(* IEC 61131-3 sources: iecf/harness/cases, 218 files *)

(* ---- autoaddrsections.st ---- *)
(* TwinCAT's `*` structures where Ed.3 6.4.4.8 refuses them
   (auto-addresses, W0020), as TcOpen's TcoEthercatMasterDevice: a
   block's VAR_INPUT, placed per instance as a VAR's, and a method's
   VAR, plain memory of the call; and its VAR_OUTPUT, which Ed.3
   allows, placed per instance.
   Placed by path, nothing stated: M: P.M.INPUTS.A 0, P.SRC.A 2.
   Q: P.M.INPUTS.B 0, P.M.OUTPUTS.Q 2, P.SRC.B 4.
   Worked by hand, k counting 1, 2: src.a := k, src.b := k * 10; the
   call m(Inputs := src) writes m.Inputs' places; Sum copies Inputs into
   its own copy, adds 100 to the copy's a (not the image's), gives
   a + b to Outputs.q.
   Tick 0: Q 10, 111, 10; M 1, 1. Tick 1: Q 20, 122, 20; M 2, 2.
   reference-skip: not IEC 61131-3. *)
TYPE Io : STRUCT
  a AT %M* : INT;
  b AT %Q* : INT;
END_STRUCT;
END_TYPE
TYPE Out : STRUCT
  q AT %Q* : INT;
END_STRUCT;
END_TYPE

FUNCTION_BLOCK Master
  VAR_INPUT Inputs : Io; END_VAR
  VAR_OUTPUT Outputs : Out; END_VAR
  METHOD Sum : INT
    VAR copy : Io; END_VAR
    copy := Inputs;
    copy.a := copy.a + 100;
    Sum := copy.a + copy.b;
  END_METHOD
  Outputs.q := THIS.Sum();
END_FUNCTION_BLOCK

PROGRAM main
  VAR k : INT; src : Io; m : Master; END_VAR
  k := k + 1;
  src.a := k;
  src.b := k * 10;
  m(Inputs := src);
END_PROGRAM

CONFIGURATION cf
  RESOURCE rs ON x
    TASK tk(INTERVAL := T#10ms, PRIORITY := 1);
    PROGRAM p WITH tk : main;
  END_RESOURCE
END_CONFIGURATION

(* ---- blockdata.st ---- *)
(* A FUNCTION_BLOCK's inputs and outputs of an array, structure or
   STRING type: copied in by the call, copied out by `=>`, read from
   outside as f.hist[0] and f.text. Each tick the input %IW0 feeds an
   array and a structure; the block keeps a history of its sums. *)
TYPE
  pair : STRUCT a : INT; b : INT; END_STRUCT;
  three : ARRAY[1..3] OF INT;
  last3 : ARRAY[0..2] OF INT;
END_TYPE

FUNCTION_BLOCK acc
VAR_INPUT
  xs : three;
  p : pair;
  tag : STRING;
END_VAR
VAR_OUTPUT
  hist : last3;
  sum : INT;
  q : pair;
  text : STRING;
END_VAR
sum := xs[1] + xs[2] + xs[3];
hist[0] := hist[1];
hist[1] := hist[2];
hist[2] := sum;
q.a := p.b;
q.b := p.a;
text := CONCAT(tag, '!');
END_FUNCTION_BLOCK

PROGRAM main
VAR
  v AT %IW0 : INT;
  r_sum AT %MW0 : INT;
  r_h2 AT %MW2 : INT;
  r_h0 AT %MW4 : INT;
  r_qa AT %MW6 : INT;
  r_qb AT %MW8 : INT;
  r_len AT %MW10 : INT;
  r_same AT %MX12.0 : BOOL;
END_VAR
VAR
  xs : three;
  pr : pair;
  h : last3;
  qq : pair;
  lab : STRING;
  f : acc;
END_VAR
xs[1] := v;
xs[2] := v * 2;
xs[3] := 1;
pr.a := v;
pr.b := 5;
f(xs := xs, p := pr, tag := 'ab', hist => h, q => qq, text => lab);
r_sum := f.sum;
r_h2 := h[2];
r_h0 := f.hist[0];
r_qa := qq.a;
r_qb := qq.b;
r_len := LEN(lab);
r_same := f.text = lab;
END_PROGRAM

CONFIGURATION plant
  RESOURCE res ON PLC
    TASK fast(INTERVAL := T#10ms, PRIORITY := 0);
    PROGRAM p WITH fast : main;
  END_RESOURCE
END_CONFIGURATION

(* ---- callparts.st ---- *)
(* A part of a FUNCTION's result read where the call is: a field, an
   element, a variable of an instance (Ed.3 6.6.2.3: a call is an operand,
   and what it gives is of the result's type).
   MKP gives a PT with x = v and y[2] = v + 1; MKA an array with [1] = v
   and [3] = 2 * v; MKC a CntT called once with inc := v, so n = v. BUMP
   adds 1 to its in-out and gives a PT with x the new value.
   Worked by hand, k %IB0 1, 2, 3; j is 2:
   MKP(k).x 1, 2, 3 (%QB0). MKP(k).y[2] 2, 3, 4 (%QB1); MKP(k).y[j], the
   index computed, the same (%QB2).
   MKA(k)[3] 2, 4, 6 (%QB3). MKA(k)[k]: [1] 1, [2] 0, [3] 6 (%QB4).
   MKC(k).n 1, 2, 3 (%QB5).
   Two calls in one expression: MKP(k).x + MKA(k)[1] 2, 4, 6 (%QB6).
   In a condition: MKP(k).x > MKC(2).n only at k 3: 0, 0, 1 (%QB7).
   A call with effects is made once though a part of it is read:
   BUMP(cnt).x 1, 2, 3 (%QB8) and cnt after it 1, 2, 3 (%QB9).
   %QB10 := MKA(k)[k + 1]: [2] 0, [3] 4; at tick 2 the index is 4,
   outside 1..3: a fault (index), the statement stopped, %QB10 kept 4.
   reference-skip: the reference compiler refuses an array or an
   instance as a FUNCTION's result, and a part of a call, MKP(k).x. *)
TYPE PT : STRUCT x : INT; y : ARRAY [1..3] OF INT; END_STRUCT; END_TYPE
FUNCTION_BLOCK CntT
  VAR_INPUT inc : INT := 1; END_VAR
  VAR_OUTPUT n : INT; END_VAR
  n := n + inc;
END_FUNCTION_BLOCK
FUNCTION MKP : PT
  VAR_INPUT v : INT; END_VAR
  MKP.x := v;
  MKP.y[2] := v + 1;
END_FUNCTION
FUNCTION MKA : ARRAY [1..3] OF INT
  VAR_INPUT v : INT; END_VAR
  MKA[1] := v;
  MKA[3] := v * 2;
END_FUNCTION
FUNCTION MKC : CntT
  VAR_INPUT v : INT; END_VAR
  MKC(inc := v);
END_FUNCTION
FUNCTION BUMP : PT
  VAR_IN_OUT n : INT; END_VAR
  n := n + 1;
  BUMP.x := n;
END_FUNCTION
CONFIGURATION c
  RESOURCE r ON PLC
    TASK t(INTERVAL := T#10ms, PRIORITY := 1);
    PROGRAM p WITH t : main;
  END_RESOURCE
END_CONFIGURATION
PROGRAM main
  VAR j : INT := 2; cnt : INT; END_VAR
  VAR k AT %IB0 : SINT; END_VAR
  VAR
    q0 AT %QB0 : SINT;
    q1 AT %QB1 : SINT;
    q2 AT %QB2 : SINT;
    q3 AT %QB3 : SINT;
    q4 AT %QB4 : SINT;
    q5 AT %QB5 : SINT;
    q6 AT %QB6 : SINT;
    q7 AT %QB7 : SINT;
    q8 AT %QB8 : SINT;
    q9 AT %QB9 : SINT;
    q10 AT %QB10 : SINT;
  END_VAR
  q0 := INT_TO_SINT(MKP(k).x);
  q1 := INT_TO_SINT(MKP(k).y[2]);
  q2 := INT_TO_SINT(MKP(k).y[j]);
  q3 := INT_TO_SINT(MKA(k)[3]);
  q4 := INT_TO_SINT(MKA(k)[k]);
  q5 := INT_TO_SINT(MKC(k).n);
  q6 := INT_TO_SINT(MKP(k).x + MKA(k)[1]);
  IF MKP(k).x > MKC(2).n THEN
    q7 := 1;
  ELSE
    q7 := 0;
  END_IF;
  q8 := INT_TO_SINT(BUMP(cnt).x);
  q9 := INT_TO_SINT(cnt);
  q10 := INT_TO_SINT(MKA(k)[k + 1]);
END_PROGRAM

(* ---- chars.st ---- *)
(* CHAR (Ed.3 Table 10, a Latin-1 character in iecf, docs/dependencies.md):
   CHAR#'X', CHAR#16#41 and an untyped 'X' where a CHAR is wanted (Table
   6, 1b); at an address, in an array and a structure, an initial value,
   a function block's input and output, a function's input and result;
   compared, MAX, SEL; CHAR_TO_BYTE and BYTE_TO_CHAR (binary transfer,
   Table 25), CHAR_TO_USINT; to a STRING, implicitly and by
   CHAR_TO_STRING, and in CONCAT; FIND of a CHAR in a STRING (Table 34,
   NOTE 3); STRING_TO_CHAR, the first character - an empty string gives
   '$00', flagged CONVERSION.
   Worked by hand: tick 0, bin 16#62 ('b'): qc 'b' (16#62), qn 16#63,
   qa 'A' (16#41), qm 'b', qlt TRUE, qeq TRUE, qs 'xb', qf 'x', qu 98,
   qp 21 (FIND(s, c) 2, FIND(s, CHAR#'x') 1).
   Tick 1, bin 16#30 ('0'): qc '0', qn '1', qm 'b' (MAX of '0' and 'b'),
   qlt TRUE, qeq FALSE, qs 'x0', qf 'x', qu 48, qp 21; then the empty string,
   flag CONVERSION.
   reference-skip: CHAR is Ed.3's; the reference compiler (Ed.2) has none. *)
TYPE rec : STRUCT c : CHAR := 'z'; n : USINT; END_STRUCT; END_TYPE

FUNCTION next_char : CHAR
VAR_INPUT c : CHAR; END_VAR
next_char := BYTE_TO_CHAR(USINT_TO_BYTE(CHAR_TO_USINT(c) + 1));
END_FUNCTION

FUNCTION_BLOCK keep
VAR_INPUT c : CHAR; END_VAR
VAR_OUTPUT last : CHAR := CHAR#'?'; END_VAR
last := c;
END_FUNCTION_BLOCK

PROGRAM main
VAR
  bin AT %IB0 : BYTE;
  qc AT %QB0 : CHAR;
  qn AT %QB1 : CHAR;
  qa AT %QB2 : CHAR;
  qm AT %QB3 : CHAR;
  qlt AT %QX4.0 : BOOL;
  qeq AT %QX4.1 : BOOL;
  qu AT %QB5 : USINT;
  qs AT %QB6 : STRING[3];
  qf AT %QB10 : CHAR;
  qp AT %QB11 : SINT;
END_VAR
VAR
  c : CHAR;
  arr : ARRAY[0..1] OF CHAR := [CHAR#'b', 'a'];
  r : rec;
  k : keep;
  s : STRING[3];
  e : STRING[3] := '';
END_VAR
c := BYTE_TO_CHAR(bin);
qc := c;
qn := next_char(c);
qa := CHAR#16#41;
qm := MAX(c, arr[0]);
qlt := c < r.c;
qeq := c = 'b';
k(c := c);
s := CONCAT('x', k.last);
qs := s;
qf := STRING_TO_CHAR(s);
qp := INT_TO_SINT(FIND(s, c) * 10 + FIND(IN1 := s, IN2 := CHAR#'x'));
qu := CHAR_TO_USINT(SEL(TRUE, arr[1], c));
qu := CHAR_TO_USINT(c);
IF c = '0' THEN
  qf := STRING_TO_CHAR(e);
END_IF;
END_PROGRAM

CONFIGURATION Plant
  RESOURCE r ON PLC
    TASK fast(INTERVAL := T#10ms, PRIORITY := 1);
    PROGRAM p WITH fast : main;
  END_RESOURCE
END_CONFIGURATION

(* ---- codesysabstract.st ---- *)
(* An ABSTRACT function block with no ABSTRACT method (codesys-oo), as
   TcOpen's TcoObject and TcoStateBase: ABSTRACT says only that it has
   no instances. Base's Run and Name are implemented; Job EXTENDS Base,
   overrides Name, and is reached through a REFERENCE TO Base, its
   override dynamically bound.
   Worked by hand, each tick: j.count + 1 through Base's Run, Name of
   Job 7 (Base's would be 1). Tick 1: 1, 7; tick 2: 2, 7.
   reference-skip: not IEC 61131-3. *)
FUNCTION_BLOCK ABSTRACT Base
  VAR_OUTPUT count : INT; END_VAR
  METHOD Run
    count := count + 1;
  END_METHOD
  METHOD Name : INT
    Name := 1;
  END_METHOD
END_FUNCTION_BLOCK

FUNCTION_BLOCK Job EXTENDS Base
  METHOD Name : INT
    Name := 7;
  END_METHOD
END_FUNCTION_BLOCK

PROGRAM main
  VAR j : Job; r : REFERENCE TO Base; END_VAR
  VAR q0 AT %QW0 : INT; q2 AT %QW2 : INT; END_VAR
  r REF= j;
  r.Run();
  q0 := j.count;
  q2 := r.Name();
END_PROGRAM

CONFIGURATION cf
  RESOURCE r ON x
    TASK tk(INTERVAL := T#10ms, PRIORITY := 1);
    PROGRAM p WITH tk : main;
  END_RESOURCE
END_CONFIGURATION

(* ---- codesysactioncall.st ---- *)
(* CODESYS's and TwinCAT's direct call of an ACTION (action-call):
   counter's own tick, which s0 runs every scan (N, never leaving it),
   calls inc bare; main calls inc too, through the instance, from
   outside. Neither call is tick's: a step runs that one, and a direct
   call of it is refused (crates/iecf-sema/tests/check.rs).
   Worked by hand: each tick, c() runs tick (+1) then main calls
   inc() itself (+1): n grows by 2 a tick, q := c.n after both.
   %QW0: tick 0 q 2, tick 1 q 4, tick 2 q 6.
   reference-skip: not IEC 61131-3. *)
FUNCTION_BLOCK counter
  VAR_OUTPUT n : INT; END_VAR
  INITIAL_STEP s0 : tick(N); END_STEP
  TRANSITION FROM s0 TO s0 := FALSE; END_TRANSITION
  ACTION tick : inc(); END_ACTION
  ACTION inc : n := n + 1; END_ACTION
END_FUNCTION_BLOCK

PROGRAM main
  VAR c : counter; END_VAR
  VAR q AT %QW0 : INT; END_VAR
  c();
  c.inc();
  q := c.n;
END_PROGRAM

CONFIGURATION cf
  RESOURCE r ON x
    TASK tk(INTERVAL := T#10ms, PRIORITY := 1);
    PROGRAM p WITH tk : main;
  END_RESOURCE
END_CONFIGURATION

(* ---- codesysaddedinout.st ---- *)
(* A derived block that adds an in-out, standing where its base is
   wanted (codesys-oo), as TcOpen's TcoCylinderMoveTask, which adds
   MoveToPositionSignal to TcoTask and is given as `refInverseTask :
   REFERENCE TO TcoTask`. A call through the base binds only the
   base's; the added in-out keeps what the last call bound, and one
   never bound is a NULL fault where the body uses it.
   Worked by hand: tick 1, m1(sig := a) sets a TRUE (from FALSE),
   then r REF= m1, r() through Job: sig still a, set FALSE; runs 2.
   Tick 2: the same, a TRUE then FALSE, runs 4; then go := TRUE.
   Tick 3: as tick 2, runs 6, then r REF= m2, never called: r.Count()
   is a method, 1; r() reaches Mover's body, `sig := NOT sig` on an
   in-out never bound: fault NULL, main line 39.
   reference-skip: not IEC 61131-3 (Ed.3 6.6.8.4 refuses it). *)
FUNCTION_BLOCK Job
  VAR_OUTPUT runs : INT; END_VAR
  METHOD Count : INT
    Count := 1;
  END_METHOD
  runs := runs + 1;
END_FUNCTION_BLOCK

FUNCTION_BLOCK Mover EXTENDS Job
  VAR_IN_OUT sig : BOOL; END_VAR
  SUPER^();
  sig := NOT sig;
END_FUNCTION_BLOCK

PROGRAM main
  VAR m1 : Mover; m2 : Mover; r : REFERENCE TO Job; a : BOOL; go : BOOL; n : INT; END_VAR
  VAR q0 AT %QX0.0 : BOOL; q2 AT %QW2 : INT; q4 AT %QW4 : INT; END_VAR
  m1(sig := a);
  r REF= m1;
  r();
  q0 := a;
  q2 := m1.runs;
  IF go THEN
    r REF= m2;
    q4 := r.Count();
    r();
  END_IF
  go := m1.runs >= 4;
END_PROGRAM

CONFIGURATION cf
  RESOURCE r ON x
    TASK tk(INTERVAL := T#10ms, PRIORITY := 1);
    PROGRAM p WITH tk : main;
  END_RESOURCE
END_CONFIGURATION

(* ---- codesysany.st ---- *)
(* ANY as an input (any-input), as CODESYS passes one and TcOpen's
   StringBuilder reads it: its type class, a pointer to the value, its
   size. Worked by hand:
   %QW0 Kind(i), an INT 7: read through the pointer, 7 + 1000 = 1007;
   %QW2 Kind(r), a REAL: 2; %QW4 Kind(5), a literal, an INT: 1005;
   %QW6 b.Add(i) adds through its pointer: i 7 -> 8, b's own total 8;
   %QW8 Kind(s), a STRING(20): neither, its size, 21 bytes.
   %QW10 a block's input: Sz(Data := r), a REAL's 4 bytes.
   cycle 1: i 8: 1008, 2, 1005, total 8 + 9 = 17 (i 9), 21, 4.
   reference-skip: not IEC 61131-3. *)
FUNCTION Kind : INT
VAR_INPUT Data : ANY; END_VAR
VAR p : POINTER TO INT; END_VAR
IF Data.TypeClass = __SYSTEM.TYPE_CLASS.TYPE_INT THEN
  p := Data.pValue;
  Kind := p^ + 1000;
ELSIF Data.TypeClass = __SYSTEM.TYPE_CLASS.TYPE_REAL THEN
  Kind := 2;
ELSE
  Kind := DINT_TO_INT(Data.diSize);
END_IF
END_FUNCTION

FUNCTION_BLOCK Acc
VAR_OUTPUT total : INT; END_VAR
METHOD PUBLIC Add : INT
VAR_INPUT Data : ANY; END_VAR
VAR p : POINTER TO INT; c : __SYSTEM.TYPE_CLASS; END_VAR
c := Data.TypeClass;
IF c = __SYSTEM.TYPE_CLASS.TYPE_INT THEN
  p := Data.pValue;
  p^ := p^ + 1;
  total := total + p^;
END_IF
Add := total;
END_METHOD
END_FUNCTION_BLOCK

FUNCTION_BLOCK Sz
VAR_INPUT Data : ANY; END_VAR
VAR_OUTPUT n : INT; END_VAR
n := DINT_TO_INT(Data.diSize);
END_FUNCTION_BLOCK

PROGRAM main
  VAR i : INT := 7; r : REAL; s : STRING(20); b : Acc; t : INT; z4 : Sz; END_VAR
  VAR x AT %QW0 : INT; y AT %QW2 : INT; z AT %QW4 : INT; w AT %QW6 : INT; v AT %QW8 : INT; u AT %QW10 : INT; END_VAR
  x := Kind(i);
  y := Kind(Data := r);
  z := Kind(5);
  t := b.Add(i);
  w := b.total;
  v := Kind(s);
  z4(Data := r);
  u := z4.n;
END_PROGRAM

CONFIGURATION cf
  RESOURCE r ON x
    TASK tk(INTERVAL := T#10ms, PRIORITY := 1);
    PROGRAM p WITH tk : main;
  END_RESOURCE
END_CONFIGURATION

(* ---- codesysargs.st ---- *)
(* Found in OSCAT NETWORK and BUILDING: a call's arguments in order
   first, then by name (mixed-arguments). Worked by hand:
   %QW0: F(1, c := 3, b := 2): a 1, b 2, c 3: 123.
   %QW2: F(1, 2, c := 4, o => s): 124, and s := 1 + 2 + 4 = 7 (%QW4).
   %QW6: sum(5, y := 6), then sum.s: 5 + 6 = 11.
   %QW8: LIMIT(0, MX := 10, IN := 15): MN 0, the rest by name: 10.
   %QW10: sum.m(9, v := 2), a method: 9 - 2 = 7.
   reference-skip: not IEC 61131-3. *)
FUNCTION F : INT
  VAR_INPUT a : INT; b : INT; c : INT; END_VAR
  VAR_OUTPUT o : INT; END_VAR
  F := a * 100 + b * 10 + c;
  o := a + b + c;
END_FUNCTION

FUNCTION_BLOCK ACC
  VAR_INPUT x : INT; y : INT; END_VAR
  VAR_OUTPUT s : INT; END_VAR
  METHOD PUBLIC m : INT
    VAR_INPUT u : INT; v : INT; END_VAR
    m := u - v;
  END_METHOD
  s := x + y;
END_FUNCTION_BLOCK

PROGRAM main
  VAR sum : ACC; END_VAR
  VAR
    q0 AT %QW0 : INT; q1 AT %QW2 : INT; s AT %QW4 : INT; q3 AT %QW6 : INT;
    q4 AT %QW8 : INT; q5 AT %QW10 : INT;
  END_VAR
  q0 := F(1, c := 3, b := 2);
  q1 := F(1, 2, c := 4, o => s);
  sum(5, y := 6);
  q3 := sum.s;
  q4 := LIMIT(0, MX := 10, IN := 15);
  q5 := sum.m(9, v := 2);
END_PROGRAM

CONFIGURATION cf
  RESOURCE r ON x
    TASK tk(INTERVAL := T#10ms, PRIORITY := 1);
    PROGRAM p WITH tk : main;
  END_RESOURCE
END_CONFIGURATION

(* ---- codesysbit.st ---- *)
(* CODESYS's and TwinCAT's BIT (bit): a structure's BITs packed into
   bytes from bit 0 up, a member of another type at the next whole byte
   aligned to its size; a function block's BIT a BOOL. Worked by hand:
   S: a %X0.0, b %X0.1, c %X0.2, n %B2 (INT, aligned to 2), d %X4.0.
   a, c and d set, n := 5: its bytes, read through V's raw,
   %QB0..4 05 00 05 00 01.
   un.d := 16#00000105: byte 0 is 2#101, byte 1 is 1.
   %QB5 bits[0].b0 01, %QB6 bits[0].b2 01, %QB7 bits[1].b0 01,
   %QB8 bits[0].b1 00, %QB9 one (a BIT in a UNION, bit 0) 01,
   %QB10 f.y, NOT bits[0].b1, 01; %QB11 00.
   un.bits[3].b7 := TRUE sets the DWORD's top bit:
   %QD12 16#80000105, 05 01 00 80.
   reference-skip: not IEC 61131-3. *)
TYPE
  S : STRUCT
    a : BIT;
    b, c : BIT;
    n : INT;
    d : BIT;
  END_STRUCT;
  V : UNION
    s : S;
    raw : ARRAY[0..4] OF BYTE;
  END_UNION;
  B8 : STRUCT
    b0 : BIT; b1 : BIT; b2 : BIT; b3 : BIT;
    b4 : BIT; b5 : BIT; b6 : BIT; b7 : BIT;
  END_STRUCT;
  U : UNION
    d : DWORD;
    bits : ARRAY[0..3] OF B8;
    one : BIT;
  END_UNION;
END_TYPE

FUNCTION_BLOCK F
  VAR_INPUT x : BIT; END_VAR
  VAR_OUTPUT y : BOOL; END_VAR
  y := NOT x;
END_FUNCTION_BLOCK

PROGRAM main
  VAR v : V; un : U; f : F; END_VAR
  VAR
    q0 AT %QB0 : BYTE; q1 AT %QB1 : BYTE; q2 AT %QB2 : BYTE; q3 AT %QB3 : BYTE;
    q4 AT %QB4 : BYTE; q5 AT %QB5 : BYTE; q6 AT %QB6 : BYTE; q7 AT %QB7 : BYTE;
    q8 AT %QB8 : BYTE; q9 AT %QB9 : BYTE; q10 AT %QB10 : BYTE; qd AT %QD12 : DWORD;
  END_VAR
  v.s.a := TRUE;
  v.s.c := TRUE;
  v.s.n := 5;
  v.s.d := TRUE;
  q0 := v.raw[0]; q1 := v.raw[1]; q2 := v.raw[2]; q3 := v.raw[3]; q4 := v.raw[4];
  un.d := 16#00000105;
  q5 := BOOL_TO_BYTE(un.bits[0].b0);
  q6 := BOOL_TO_BYTE(un.bits[0].b2);
  q7 := BOOL_TO_BYTE(un.bits[1].b0);
  q8 := BOOL_TO_BYTE(un.bits[0].b1);
  q9 := BOOL_TO_BYTE(un.one);
  f(x := un.bits[0].b1);
  q10 := BOOL_TO_BYTE(f.y);
  un.bits[3].b7 := TRUE;
  qd := un.d;
END_PROGRAM

CONFIGURATION cf
  RESOURCE r ON x
    TASK tk(INTERVAL := T#10ms, PRIORITY := 1);
    PROGRAM p WITH tk : main;
  END_RESOURCE
END_CONFIGURATION

(* ---- codesysemptyargs.st ---- *)
(* CODESYS's and TwinCAT's empty arguments (empty-arguments): a
   parameter named and given nothing, `x :=,` or `y =>,`, as their
   input assistant writes every one; TcOpen's EtherCAT calls do. It is
   left out: an instance's input keeps what it had, an output is not
   read, a FUNCTION's input is its initial value.
   Worked by hand: c.n grows by inc each call, en TRUE.
   tick 0: c(inc := 2, en :=,...): n 2, x 2; c(inc :=, ...): inc
   still 2, n 4, y 4; add3(a := 1, b :=): 1 + 10 = 11.
   A last `,` before `)` is one with no name, as TcOpen's WpfContext
   writes `outHopper => ..., );`: d(inc := 3, n => v, ) gives v 3,
   then 6; add3(a := 2, ) 12.
   tick 1: x 6, y 8, z 11.
   reference-skip: not IEC 61131-3. *)
FUNCTION_BLOCK Cnt
  VAR_INPUT inc : INT := 1; en : BOOL := TRUE; END_VAR
  VAR_OUTPUT n : INT; busy : BOOL; END_VAR
  IF en THEN n := n + inc; END_IF;
  busy := n > 5;
END_FUNCTION_BLOCK

FUNCTION add3 : INT
  VAR_INPUT a : INT; b : INT := 10; END_VAR
  add3 := a + b;
END_FUNCTION

PROGRAM main
  VAR c : Cnt; d : Cnt; END_VAR
  VAR x AT %QB0 : SINT; y AT %QB1 : SINT; z AT %QB2 : SINT; v AT %QB3 : SINT; w AT %QB4 : SINT; END_VAR
  c(inc := 2, en :=, busy =>, n => x);
  c(inc :=,
    en :=,
    busy =>,
    n => y);
  z := TO_SINT(add3(a := 1, b :=));
  d(inc := 3,
    n => v,
   );
  w := TO_SINT(add3(a := 2, ));
END_PROGRAM

CONFIGURATION cf
  RESOURCE r ON x
    TASK tk(INTERVAL := T#10ms, PRIORITY := 1);
    PROGRAM p WITH tk : main;
  END_RESOURCE
END_CONFIGURATION

(* ---- codesysexprstmt.st ---- *)
(* An expression standing as a statement (expression-statements), as
   TcOpen's tests read a property for what its GET does,
   `_sutNotInitialized.IsTrue;`, `_sut_A.Invoke().Done;`: every call in
   it made, its value unused; one with no call does nothing.
   Worked by hand, each tick: s.IsTrue's GET counts 1; t.Invoke() 1 and
   Done's GET 1, through the interface Invoke gives; Bump(n := k) + 1
   adds 1 to k (from 10); s.flag and arr[i], i out of bounds, nothing.
   Tick 1: 1, 1, 1, 11; tick 2: 2, 2, 2, 12.
   IT's GET holds an empty VAR ... END_VAR, as TwinCAT writes one
   (properties).
   reference-skip: not IEC 61131-3. *)
INTERFACE IT
  PROPERTY Done : BOOL
    GET
    VAR
    END_VAR
    END_GET
  END_PROPERTY
END_INTERFACE

FUNCTION_BLOCK Sig
  VAR_OUTPUT gets : INT; flag : BOOL; END_VAR
  PROPERTY IsTrue : BOOL
    GET
      gets := gets + 1;
      IsTrue := flag;
    END_GET
  END_PROPERTY
END_FUNCTION_BLOCK

FUNCTION_BLOCK Job IMPLEMENTS IT
  VAR_OUTPUT invokes : INT; dones : INT; END_VAR
  METHOD Invoke : IT
    invokes := invokes + 1;
    Invoke := THIS^;
  END_METHOD
  PROPERTY Done : BOOL
    GET
      dones := dones + 1;
      Done := TRUE;
    END_GET
  END_PROPERTY
END_FUNCTION_BLOCK

FUNCTION Bump : INT
  VAR_IN_OUT n : INT; END_VAR
  n := n + 1;
  Bump := n;
END_FUNCTION

PROGRAM main
  VAR s : Sig; t : Job; k : INT := 10; arr : ARRAY[1..2] OF INT; i : INT := 5; END_VAR
  VAR q0 AT %QW0 : INT; q2 AT %QW2 : INT; q4 AT %QW4 : INT; q6 AT %QW6 : INT; END_VAR
  s.IsTrue;
  t.Invoke().Done;
  Bump(n := k) + 1;
  s.flag;
  arr[i];
  q0 := s.gets;
  q2 := t.invokes;
  q4 := t.dones;
  q6 := k;
END_PROGRAM

CONFIGURATION cf
  RESOURCE r ON x
    TASK tk(INTERVAL := T#10ms, PRIORITY := 1);
    PROGRAM p WITH tk : main;
  END_RESOURCE
END_CONFIGURATION

(* ---- codesysfbinit.st ---- *)
(* CODESYS's FB_init (fb-init), as TcOpen gives it: `child : T(THIS^,
   eMode.Keep)`. Worked by hand, at the cold start:
   %QW0: Base's FB_init, then Derived's, each its own: order 1 * 10 + 2,
   12.
   %QW2: the parent given, THIS^, Root: its Depth, 7.
   %QW4: the mode given, eMode.Keep, 1.
   %QX6.0: bInitRetains at a cold start: TRUE.
   %QW8: Counter's FB_init, the two flags alone, called once: 1.
   %QW10: Wider, derived from Derived, its FB_init naming the two
   inputs it shares p and m and adding level: Base's, Derived's and
   its own, 123; %QW12 level, 42; %QW14 Base's mode, given by place
   to each, 1.
   reference-skip: not IEC 61131-3. *)
INTERFACE IObject
  METHOD Depth : INT
  END_METHOD
END_INTERFACE

TYPE eMode : (None, Keep); END_TYPE

FUNCTION_BLOCK Base
  VAR _parent : IObject; _mode : eMode; order : INT; cold : BOOL; END_VAR
  METHOD FB_init : BOOL
    VAR_INPUT bInitRetains : BOOL; bInCopyCode : BOOL; parent : IObject; mode : eMode; END_VAR
    _parent := parent;
    _mode := mode;
    order := order * 10 + 1;
    cold := bInitRetains;
  END_METHOD
  METHOD ParentDepth : INT
    ParentDepth := _parent.Depth();
  END_METHOD
END_FUNCTION_BLOCK

FUNCTION_BLOCK Derived EXTENDS Base
  METHOD FB_init : BOOL
    VAR_INPUT bInitRetains : BOOL; bInCopyCode : BOOL; parent : IObject; mode : eMode; END_VAR
    order := order * 10 + 2;
  END_METHOD
END_FUNCTION_BLOCK

FUNCTION_BLOCK Counter
  VAR_OUTPUT n : INT; END_VAR
  METHOD FB_init : BOOL
    VAR_INPUT bInitRetains : BOOL; bInCopyCode : BOOL; END_VAR
    n := n + 1;
  END_METHOD
END_FUNCTION_BLOCK

FUNCTION_BLOCK Wider EXTENDS Derived
  VAR extra : INT; END_VAR
  METHOD FB_init : BOOL
    VAR_INPUT bInitRetains : BOOL; bInCopyCode : BOOL; p : IObject; m : eMode; level : INT; END_VAR
    extra := level;
    order := order * 10 + 3;
  END_METHOD
END_FUNCTION_BLOCK

FUNCTION_BLOCK Root IMPLEMENTS IObject
  VAR child : Derived(THIS^, eMode.Keep); END_VAR
  VAR wide : Wider(THIS^, eMode.Keep, 42); END_VAR
  METHOD Depth : INT
    Depth := 7;
  END_METHOD
END_FUNCTION_BLOCK

PROGRAM main
  VAR r : Root; plain : Counter; END_VAR
  VAR q0 AT %QW0 : INT; q1 AT %QW2 : INT; q2 AT %QW4 : INT; q3 AT %QX6.0 : BOOL; q4 AT %QW8 : INT;
      q5 AT %QW10 : INT; q6 AT %QW12 : INT; q7 AT %QW14 : INT; END_VAR
  q0 := r.child.order;
  q1 := r.child.ParentDepth();
  q2 := TO_INT(r.child._mode);
  q3 := r.child.cold;
  q4 := plain.n;
  q5 := r.wide.order;
  q6 := r.wide.extra;
  q7 := TO_INT(r.wide._mode);
END_PROGRAM

CONFIGURATION cf
  RESOURCE r ON x
    TASK tk(INTERVAL := T#10ms, PRIORITY := 1);
    PROGRAM p WITH tk : main;
  END_RESOURCE
END_CONFIGURATION

(* ---- codesyshdrsemi.st ---- *)
(* A `;` closing a header before its declarations (header-semicolon),
   as TcOpen's TcoInsight writes `METHOD SetUserDataAsByte : BOOL;`, and
   a method's variable named as its block's (shadowing), hiding it in
   the method, THIS^.n still the block's.
   Worked by hand, each tick: b(n := 100) sets the block's n, hits + 1;
   b.Add(n := 5) adds its own n, 5, to total and 1 to the block's n,
   101; b.Peek() reads the block's n, 101; F(a := 21) 42.
   Tick 1: Add 5, Peek 101, b.n 101, hits 1, F 42.
   Tick 2: Add 10, Peek 101, b.n 101, hits 2, F 42.
   reference-skip: not IEC 61131-3. *)
FUNCTION F : INT;
  VAR_INPUT a : INT; END_VAR
  F := a * 2;
END_FUNCTION

FUNCTION_BLOCK Blk
  VAR_INPUT n : INT; END_VAR
  VAR_OUTPUT hits : INT; END_VAR
  VAR total : INT; END_VAR
  METHOD Add : INT;
    VAR_INPUT n : INT; END_VAR
    total := total + n;
    THIS^.n := THIS^.n + 1;
    Add := total;
  END_METHOD
  METHOD Peek : INT;
    Peek := n;
  END_METHOD
  hits := hits + 1;
END_FUNCTION_BLOCK

PROGRAM main
  VAR b : Blk; END_VAR
  VAR q0 AT %QW0 : INT; q2 AT %QW2 : INT; q4 AT %QW4 : INT; q6 AT %QW6 : INT; q8 AT %QW8 : INT; END_VAR
  b(n := 100);
  q0 := b.Add(n := 5);
  q2 := b.Peek();
  q4 := b.n;
  q6 := b.hits;
  q8 := F(a := 21);
END_PROGRAM

CONFIGURATION cf
  RESOURCE r ON x
    TASK tk(INTERVAL := T#10ms, PRIORITY := 1);
    PROGRAM p WITH tk : main;
  END_RESOURCE
END_CONFIGURATION

(* ---- codesysinout.st ---- *)
(* A method using its block's VAR_IN_OUT (method-in-outs), as TcOpen's
   do, CODESYS warning C0371: what the block's last call bound.
   Worked by hand:
   %QW0, %QW2: d1 := 5, d2 := 6; ax(drive := d1), ax.Stop() sets d1 to 0;
   ax(drive := d2), ax.Stop() sets d2 to 0: 0 and 0.
   %QW4: p.speed through the structure in-out: Stop writes 7.
   %QW6: set to 1 before bx.Stop(), bx never called: NULL fault on the
   line of bx.Stop() (34), the task stops there; q3 stays 1.
   reference-skip: not IEC 61131-3. *)
TYPE Info : STRUCT speed : INT; END_STRUCT; END_TYPE

FUNCTION_BLOCK Axis
  VAR_IN_OUT drive : INT; data : Info; END_VAR
  METHOD PUBLIC Stop
    drive := 0;
    data.speed := 7;
  END_METHOD
  drive := drive;
END_FUNCTION_BLOCK

PROGRAM main
  VAR ax : Axis; bx : Axis; d1 : INT := 5; d2 : INT := 6; p : Info; END_VAR
  VAR q0 AT %QW0 : INT; q1 AT %QW2 : INT; q2 AT %QW4 : INT; q3 AT %QW6 : INT; END_VAR
  ax(drive := d1, data := p);
  ax.Stop();
  ax(drive := d2, data := p);
  ax.Stop();
  q0 := d1;
  q1 := d2;
  q2 := p.speed;
  q3 := 1;

  bx.Stop();
  q3 := 2;
END_PROGRAM

CONFIGURATION cf
  RESOURCE r ON x
    TASK tk(INTERVAL := T#10ms, PRIORITY := 1);
    PROGRAM p WITH tk : main;
  END_RESOURCE
END_CONFIGURATION

(* ---- codesysinoutkept.st ---- *)
(* method-in-outs: a method's own in-out given to a block's in-out that
   a method of the block uses after the call, kept past the method's
   call; the call of the method gives a variable that lives as long as
   the program, two methods deep (Pass gives y to Run's x, Run to the
   block's v).
   Worked by hand, g 10: tick 0: u.Pass(y := g) binds t.v to g; u.Tick()
   bumps it: g 11. Ticks 1, 2, Pass not called: g 12, 13.
   %QW0 11, 12, 13.
   reference-skip: not IEC 61131-3. *)
FUNCTION_BLOCK Holder
  VAR_IN_OUT v : INT; END_VAR
  METHOD PUBLIC Bump
    v := v + 1;
  END_METHOD
END_FUNCTION_BLOCK

FUNCTION_BLOCK User
  VAR t : Holder; END_VAR
  METHOD PUBLIC Run
    VAR_IN_OUT x : INT; END_VAR
    t(v := x);
  END_METHOD
  METHOD PUBLIC Pass
    VAR_IN_OUT y : INT; END_VAR
    THIS^.Run(x := y);
  END_METHOD
  METHOD PUBLIC Tick
    t.Bump();
  END_METHOD
END_FUNCTION_BLOCK

PROGRAM main
  VAR u : User; g : INT := 10; started : BOOL; END_VAR
  VAR q0 AT %QW0 : INT; END_VAR
  IF NOT started THEN
    u.Pass(y := g);
    started := TRUE;
  END_IF
  u.Tick();
  q0 := g;
END_PROGRAM

CONFIGURATION cf
  RESOURCE r ON x
    TASK tk(INTERVAL := T#10ms, PRIORITY := 1);
    PROGRAM p WITH tk : main;
  END_RESOURCE
END_CONFIGURATION

(* ---- codesysinoutref.st ---- *)
(* method-in-outs: a method's own in-out bound by REF= to a reference
   of its block, which outlives the call, as TcOpen's
   TcoInspector.UpdateComprehensiveResult(VAR_IN_OUT inoResult) keeps
   `_refOverallResult REF= inoResult`: kept past the method's call, and
   each call of the method gives a variable that lives as long as the
   program, two methods deep (Pass gives y to Update's x).
   Worked by hand, g 1: tick 0: k.Pass(y := g) binds k.r to g;
   k.Tick() adds 5 through it: g 6. Ticks 1, 2, Pass not called: 11,
   16. %QW0 6, 11, 16.
   reference-skip: not IEC 61131-3. *)
FUNCTION_BLOCK Keeper
  VAR r : REFERENCE TO INT; END_VAR
  METHOD PUBLIC Update
    VAR_IN_OUT x : INT; END_VAR
    r REF= x;
  END_METHOD
  METHOD PUBLIC Pass
    VAR_IN_OUT y : INT; END_VAR
    THIS^.Update(x := y);
  END_METHOD
  METHOD PUBLIC Tick
    IF __ISVALIDREF(r) THEN
      r := r + 5;
    END_IF
  END_METHOD
END_FUNCTION_BLOCK

PROGRAM main
  VAR k : Keeper; g : INT := 1; started : BOOL; END_VAR
  VAR q0 AT %QW0 : INT; END_VAR
  IF NOT started THEN
    k.Pass(y := g);
    started := TRUE;
  END_IF
  k.Tick();
  q0 := g;
END_PROGRAM

CONFIGURATION cf
  RESOURCE r ON x
    TASK tk(INTERVAL := T#10ms, PRIORITY := 1);
    PROGRAM p WITH tk : main;
  END_RESOURCE
END_CONFIGURATION

(* ---- codesysinoutvalid.st ---- *)
(* A method testing its block's VAR_IN_OUT with __ISVALIDREF
   (method-in-outs), as TcOpen's tasks do before using one: FALSE until
   a call of the block binds it, and a use the test guards is no fault.
   Worked by hand, s.d from 3:
   cycle 0: i.M() before any call of i: unbound, -1 (the ELSIF that
     reads io not tested); i(io := s): d 6; i.M(): d 7, 7.
   cycle 1: i.M(): bound by the last call, d 8, 8; i(): 16; i.M(): 17.
   A derived block's body tests the in-out it inherits, bound by its
   call: %QW4 1, and its d (from 5) 5 + 10 = 15 at %QW6, 25 next.
   reference-skip: not IEC 61131-3. *)
TYPE St : STRUCT d : INT; END_STRUCT; END_TYPE

FUNCTION_BLOCK B
VAR_IN_OUT io : St; END_VAR
METHOD PUBLIC M : INT
IF NOT __ISVALIDREF(io) THEN
  M := -1;
ELSIF io.d > 1000 THEN
  M := 0;
ELSE
  THIS^.io.d := io.d + 1;
  M := io.d;
END_IF
END_METHOD
io.d := io.d * 2;
END_FUNCTION_BLOCK

FUNCTION_BLOCK D EXTENDS B
VAR_OUTPUT ok : BOOL; END_VAR
ok := __ISVALIDREF(io);
IF __ISVALIDREF(THIS^.io) THEN
  io.d := io.d + 10;
END_IF
END_FUNCTION_BLOCK

PROGRAM main
  VAR i : B; s : St := (d := 3); j : D; t : St := (d := 5); END_VAR
  VAR a AT %QW0 : INT; b AT %QW2 : INT; c AT %QW4 : INT; e AT %QW6 : INT; END_VAR
  a := i.M();
  i(io := s);
  b := i.M();
  j(io := t);
  c := BOOL_TO_INT(j.ok);
  e := t.d;
END_PROGRAM

CONFIGURATION cf
  RESOURCE r ON x
    TASK tk(INTERVAL := T#10ms, PRIORITY := 1);
    PROGRAM p WITH tk : main;
  END_RESOURCE
END_CONFIGURATION

(* ---- codesysitfspecs.st ---- *)
(* CODESYS's and TwinCAT's PUBLIC and FINAL on an interface's method
   or property (codesys-oo), as TcOpen writes `METHOD PUBLIC FINAL
   StepIn` in ITcoSequencerModeController: PUBLIC is what a prototype
   is, FINAL has no effect. Worked by hand:
   %QW0 through I, d is a D, whose Advance overrides B's although I's is
        FINAL: 2; B's Speed 5: 7.
   reference-skip: not IEC 61131-3. *)
INTERFACE I
  METHOD PUBLIC FINAL Advance : INT
  END_METHOD
  PROPERTY PUBLIC Speed : INT
  GET
  END_GET
  END_PROPERTY
END_INTERFACE
FUNCTION_BLOCK B IMPLEMENTS I
  METHOD PUBLIC Advance : INT
    Advance := 1;
  END_METHOD
  PROPERTY PUBLIC Speed : INT
  GET
    Speed := 5;
  END_GET
  END_PROPERTY
END_FUNCTION_BLOCK
FUNCTION_BLOCK D EXTENDS B
  METHOD PUBLIC Advance : INT
    Advance := 2;
  END_METHOD
END_FUNCTION_BLOCK
PROGRAM main
  VAR d : D; i : I; END_VAR
  VAR n AT %QW0 : INT; END_VAR
  i := d;
  n := i.Advance() + i.Speed;
END_PROGRAM
CONFIGURATION cf
  RESOURCE r ON x
    TASK tk(INTERVAL := T#10ms, PRIORITY := 1);
    PROGRAM p WITH tk : main;
  END_RESOURCE
END_CONFIGURATION

(* ---- codesysitftwice.st ---- *)
(* CODESYS's and TwinCAT's IMPLEMENTS naming an interface twice
   (codesys-oo), as TcOpen's TcoInputDialog writes `IMPLEMENTS
   ITcoInputDialogAnswer, ITcoInputDialogAnswer`: it counts once,
   W0019. Worked by hand:
   %QW0 through I, d is a D, whose Answer overrides B's: 2, then 4.
   reference-skip: not IEC 61131-3. *)
INTERFACE I
  METHOD Answer : INT
  END_METHOD
END_INTERFACE
FUNCTION_BLOCK B IMPLEMENTS I, I
  VAR n : INT; END_VAR
  METHOD PUBLIC Answer : INT
    n := n + 1;
    Answer := n;
  END_METHOD
END_FUNCTION_BLOCK
FUNCTION_BLOCK D EXTENDS B
  METHOD PUBLIC Answer : INT
    n := n + 2;
    Answer := n;
  END_METHOD
END_FUNCTION_BLOCK
PROGRAM main
  VAR d : D; i : I; END_VAR
  VAR q AT %QW0 : INT; END_VAR
  i := d;
  q := i.Answer();
END_PROGRAM
CONFIGURATION cf
  RESOURCE r ON x
    TASK tk(INTERVAL := T#10ms, PRIORITY := 1);
    PROGRAM p WITH tk : main;
  END_RESOURCE
END_CONFIGURATION

(* ---- codesysitfzero.st ---- *)
(* An interface compared with 0 (codesys-oo), CODESYS's test of one for
   NULL, as TcOpen tests its parent before reaching through it.
   Worked by hand:
   cycle 0: ref NULL: %QW0 (ref = 0) 1; the IF's AND_THEN calls no method
     of NULL: %QW2 0; ref := blk: %QW4 (ref <> 0) 1; %QW6 0 <> ref, 1.
   cycle 1: ref is blk's from cycle 0: %QW0 0; %QW2 blk.Get() 5; 1; 1.
   0 given to an interface (codesys-oo), its NULL: r2 starts 0, is blk
   in the cycle, and 0 again at its end. Each cycle: %QW8 (r2 = 0) 1;
   %QW10 (r2 <> 0) once r2 := blk, 1; %QW12 Has(i := 0) + 10 *
   Has(i := blk) = 0 + 10 = 10; %QW14 (Pick() = 0) 1; %QW16 r2's
   method not called once r2 := 0: 7.
   reference-skip: not IEC 61131-3. *)
INTERFACE I
METHOD Get : INT
END_METHOD
END_INTERFACE

FUNCTION Has : INT
  VAR_INPUT i : I; END_VAR
  Has := BOOL_TO_INT(i <> 0);
END_FUNCTION

FUNCTION Pick : I
  Pick := 0;
END_FUNCTION

FUNCTION_BLOCK A IMPLEMENTS I
METHOD PUBLIC Get : INT
Get := 5;
END_METHOD
END_FUNCTION_BLOCK

PROGRAM main
  VAR blk : A; ref : I; r2 : I := 0; END_VAR
  VAR x AT %QW0 : INT; y AT %QW2 : INT; z AT %QW4 : INT; w AT %QW6 : INT; END_VAR
  VAR v AT %QW8 : INT; q AT %QW10 : INT; u AT %QW12 : INT; t AT %QW14 : INT; s AT %QW16 : INT; END_VAR
  v := BOOL_TO_INT(r2 = 0);
  r2 := blk;
  q := BOOL_TO_INT(r2 <> 0);
  u := Has(i := 0) + 10 * Has(i := blk);
  t := BOOL_TO_INT(Pick() = 0);
  r2 := 0;
  s := 7;
  IF r2 <> 0 THEN
    s := r2.Get();
  END_IF;
  x := BOOL_TO_INT(ref = 0);
  y := 0;
  IF ref <> 0 AND_THEN ref.Get() > 0 THEN
    y := ref.Get();
  END_IF;
  ref := blk;
  z := BOOL_TO_INT(ref <> 0);
  w := BOOL_TO_INT(0 <> ref);
END_PROGRAM

CONFIGURATION cf
  RESOURCE r ON x
    TASK tk(INTERVAL := T#10ms, PRIORITY := 1);
    PROGRAM p WITH tk : main;
  END_RESOURCE
END_CONFIGURATION

(* ---- codesysmembershadow.st ---- *)
(* A block's members hide a library's elements of their names, as
   CODESYS's shadowing rules have it ("Local variables in the function
   block ... and in any base function blocks", "Local methods of the
   POU", before "POU or type names from a library"), as TcOpen's
   cylinders call their PROPERTY StopTask's Restore() beside
   TcoDrivesBeckhoff's FUNCTION_BLOCK StopTask. The library L
   (codesysmembershadow.d/lib.st) has a block StopTask and functions
   Helper and Twice; each 1000 or its double when reached by mistake.
   Worked by hand, each cycle:
   c (Cyl): its own PROPERTY StopTask, t's Restore() 7, %QW0 7; its own
     METHOD Helper 42, %QW2 42; L.Helper() still the library's,
     %QW4 1000; Twice(3), the library's, as nothing hides it, %QW6 6.
   d (Cyl2, from Middle, from Base): the inherited PROPERTY StopTask,
     Base's ABSTRACT one given by Middle, Restore() 7, %QW8 7; the
     inherited METHOD Helper 42, %QW10 42; an inherited variable Twice,
     an instance of T, Twice.Restore() 7, %QW12 7.
   reference-skip: not IEC 61131-3. *)
INTERFACE ITask
  METHOD Restore : INT
  END_METHOD
END_INTERFACE

FUNCTION_BLOCK T IMPLEMENTS ITask
  METHOD Restore : INT
    Restore := 7;
  END_METHOD
END_FUNCTION_BLOCK

FUNCTION_BLOCK ABSTRACT Base
  VAR t : T; Twice : T; END_VAR
  VAR_OUTPUT r1 : INT; r2 : INT; r3 : INT; r4 : INT; END_VAR
  PROPERTY ABSTRACT StopTask : ITask
    GET
    END_GET
  END_PROPERTY
  METHOD Helper : INT
    Helper := 42;
  END_METHOD
END_FUNCTION_BLOCK

FUNCTION_BLOCK Middle EXTENDS Base
  PROPERTY StopTask : ITask
    GET
      StopTask := t;
    END_GET
  END_PROPERTY
END_FUNCTION_BLOCK

FUNCTION_BLOCK Cyl
  VAR t : T; END_VAR
  VAR_OUTPUT r1 : INT; r2 : INT; r3 : INT; r4 : INT; END_VAR
  PROPERTY StopTask : ITask
    GET
      StopTask := t;
    END_GET
  END_PROPERTY
  METHOD Helper : INT
    Helper := 42;
  END_METHOD
  r1 := StopTask.Restore();
  r2 := Helper();
  r3 := L.Helper();
  r4 := Twice(3);
END_FUNCTION_BLOCK

FUNCTION_BLOCK Cyl2 EXTENDS Middle
  r1 := StopTask.Restore();
  r2 := Helper();
  r3 := Twice.Restore();
END_FUNCTION_BLOCK

PROGRAM main
  VAR c : Cyl; d : Cyl2; END_VAR
  VAR q0 AT %QW0 : INT; q1 AT %QW2 : INT; q2 AT %QW4 : INT; q3 AT %QW6 : INT;
      q4 AT %QW8 : INT; q5 AT %QW10 : INT; q6 AT %QW12 : INT; END_VAR
  c();
  d();
  q0 := c.r1; q1 := c.r2; q2 := c.r3; q3 := c.r4;
  q4 := d.r1; q5 := d.r2; q6 := d.r3;
END_PROGRAM

CONFIGURATION cf
  RESOURCE r ON x
    TASK tk(INTERVAL := T#10ms, PRIORITY := 1);
    PROGRAM p WITH tk : main;
  END_RESOURCE
END_CONFIGURATION

(* ---- codesysmix.st ---- *)
(* Two generator fixes found building the OSCAT NETWORK and BUILDING
   libraries. Worked by hand:
   %QW0: a duration times a BYTE (bit-string-arithmetic): T#100ms *
   BYTE#3 is T#300ms, as DINT 300 (BUILDING's ACTUATOR_2P).
   %QW2: inside Cron a block input named Bump shadows the FUNCTION Bump,
   which writes a global (a call with effects, so its statement is
   sequenced); arr[1] := Bump(5) calls the function: g 10 + 5 = 15, and
   g becomes 11 (NETWORK's DLOG_CRON_TAB).
   %QW4: g after the call, 11.
   reference-skip: both forms are CODESYS's, not IEC 61131-3. *)
VAR_GLOBAL g : INT := 10; END_VAR

FUNCTION Bump : INT
  VAR_INPUT x : INT; END_VAR
  VAR_EXTERNAL g : INT; END_VAR
  Bump := g + x;
  g := g + 1;
END_FUNCTION

FUNCTION_BLOCK Cron
  VAR_INPUT bump : STRING[10]; END_VAR
  VAR_OUTPUT arr : ARRAY[0..2] OF INT; END_VAR
  arr[1] := Bump(5);
END_FUNCTION_BLOCK

PROGRAM main
  VAR c : Cron; t : TIME; k : BYTE := 3; END_VAR
  VAR_EXTERNAL g : INT; END_VAR
  VAR q0 AT %QW0 : INT; q1 AT %QW2 : INT; q2 AT %QW4 : INT; END_VAR
  t := T#100ms * k;
  q0 := DINT_TO_INT(TIME_TO_DINT(t));
  c(bump := 'x');
  q1 := c.arr[1];
  q2 := g;
END_PROGRAM

CONFIGURATION cf
  RESOURCE r ON x
    TASK tk(INTERVAL := T#10ms, PRIORITY := 1);
    PROGRAM p WITH tk : main;
  END_RESOURCE
END_CONFIGURATION

(* ---- codesysnames.st ---- *)
(* Two CODESYS ways, each an extension (docs/extensions.md). Worked by
   hand:
   input-constant: Ramp's VAR_INPUT CONSTANT k is a plain input, given 3
   by the call and written in the body (k := k + 1, 4): a CONSTANT that
   means something only to CODESYS's CFC editor.
   keyword-names: step, on, r_edge and f_edge are names. step := k, 4;
   on := step + 1, 5; FOR i := 1 TO 10 BY step runs for 1, 5, 9: r_edge
   := r_edge + on three times, 15 (%QB0). f_edge := MAX(step, on), 5
   (%QB1). The SFC beside them keeps STEP as its keyword: Count's chart
   goes s0 -> s1 -> s0, its action adding 1 to n in s1, every second
   tick: after two ticks n is 1 (%QB2).
   x : BOOL R_EDGE keeps R_EDGE as its keyword: TRUE on the first tick
   only, so seen counts 1 (%QB3).
   reference-skip: neither is IEC 61131-3. *)
FUNCTION_BLOCK Ramp
  VAR_INPUT CONSTANT k : INT := 1; END_VAR
  VAR_INPUT x : BOOL R_EDGE; END_VAR
  VAR_OUTPUT r_edge, f_edge, seen : INT; END_VAR
  VAR step, on, i : INT; END_VAR
  k := k + 1;
  step := k;
  on := step + 1;
  r_edge := 0;
  FOR i := 1 TO 10 BY step DO
    r_edge := r_edge + on;
  END_FOR;
  f_edge := MAX(IN1 := step, IN2 := on);
  IF x THEN
    seen := seen + 1;
  END_IF;
END_FUNCTION_BLOCK

FUNCTION_BLOCK Count
  VAR_OUTPUT n : INT; END_VAR
  INITIAL_STEP s0 : END_STEP
  TRANSITION FROM s0 TO s1 := TRUE; END_TRANSITION
  STEP s1 : bump(P); END_STEP
  TRANSITION FROM s1 TO s0 := TRUE; END_TRANSITION
  ACTION bump : n := n + 1; END_ACTION
END_FUNCTION_BLOCK

PROGRAM main
  VAR r : Ramp; c : Count; END_VAR
  VAR
    q0 AT %QB0 : SINT;
    q1 AT %QB1 : SINT;
    q2 AT %QB2 : SINT;
    q3 AT %QB3 : SINT;
  END_VAR
  r(k := 3, x := TRUE);
  c();
  q0 := INT_TO_SINT(r.r_edge);
  q1 := INT_TO_SINT(r.f_edge);
  q2 := INT_TO_SINT(c.n);
  q3 := INT_TO_SINT(r.seen);
END_PROGRAM

CONFIGURATION cf
  RESOURCE res ON x
    TASK tk(INTERVAL := T#10ms, PRIORITY := 1);
    PROGRAM p WITH tk : main;
  END_RESOURCE
END_CONFIGURATION

(* ---- codesysobjcopy.st ---- *)
(* A block with methods used as CODESYS and TwinCAT let one be:
   declared in a method's or a FUNCTION's VAR, set up at each call
   (temp-instances), and, of its own type only, copied with := and
   given as an input (codesys-oo), as TcOpen's `_signalInfo :
   TcoSignalInfo` in a method, `_content := inoContent`, `inSignalInfo :
   TcoSignalInfo`.
   Kid EXTENDS Info and overrides Inc (+10, not +1); Info.Twice calls
   Inc through THIS^, so a Kid set up at each call must have Kid's
   methods: Twice gives 20, never 2, and starts from n = 0 each call.
   Worked by hand, each tick: Local and Fun give 20 every tick (a kept
   instance would give 40, 60); src is bumped, copied into u.inInfo by
   u(inInfo := src), bumped again, which the copy does not see, then
   copied into u.viaRef through a REFERENCE TO; u.kept := u.inInfo.
   Tick t: src.n is 2t-1 when copied in, 2t when taken by reference.
   Tick 1: 20, 20, 1, 1, 2; tick 2: 20, 20, 3, 3, 4.
   reference-skip: not IEC 61131-3. *)
FUNCTION_BLOCK Info
  VAR_OUTPUT n : INT; END_VAR
  METHOD Inc
    n := n + 1;
  END_METHOD
  METHOD Twice : INT
    THIS^.Inc();
    THIS^.Inc();
    Twice := n;
  END_METHOD
  METHOD Bump
    n := n + 1;
  END_METHOD
END_FUNCTION_BLOCK

FUNCTION_BLOCK Kid EXTENDS Info
  METHOD Inc
    n := n + 10;
  END_METHOD
END_FUNCTION_BLOCK

FUNCTION Fun : INT
  VAR k : Kid; END_VAR
  Fun := k.Twice();
END_FUNCTION

FUNCTION_BLOCK User
  VAR_INPUT inInfo : Info; END_VAR
  VAR kept : Info; viaRef : Info; END_VAR
  METHOD Local : INT
    VAR k : Kid; END_VAR
    Local := k.Twice();
  END_METHOD
  METHOD Take
    VAR_INPUT other : REFERENCE TO Info; END_VAR
    viaRef := other;
  END_METHOD
  kept := inInfo;
END_FUNCTION_BLOCK

PROGRAM main
  VAR u : User; src : Info; END_VAR
  VAR q0 AT %QW0 : INT; q2 AT %QW2 : INT; q4 AT %QW4 : INT; q6 AT %QW6 : INT; q8 AT %QW8 : INT; END_VAR
  src.Bump();
  u(inInfo := src);
  src.Bump();
  u.Take(other := src);
  q0 := u.Local();
  q2 := Fun();
  q4 := u.inInfo.n;
  q6 := u.kept.n;
  q8 := u.viaRef.n;
END_PROGRAM

CONFIGURATION cf
  RESOURCE r ON x
    TASK tk(INTERVAL := T#10ms, PRIORITY := 1);
    PROGRAM p WITH tk : main;
  END_RESOURCE
END_CONFIGURATION

(* ---- codesysoo.st ---- *)
(* CODESYS's and TwinCAT's object orientation (codesys-oo), as TcOpen
   writes it: THIS^ and SUPER^, overriding without OVERRIDE, no access
   specifier meaning PUBLIC. Worked by hand:
   %QD0: sq.Area(): side * side + SUPER^.Area(), 3.0 * 3.0 + 0.0 = 9.0,
   16#41100000.
   %QW4: sq.Describe(), Shape's, calls THIS^.Kind(): Square's override,
   2.
   %QW6: sq's body calls SUPER^(), Shape's body, once: calls = 1.
   %QW8: sq.Twice(), Shape's, calls Kind() bare, as THIS.Kind():
   Square's override, 2 * 2 = 4.
   reference-skip: not IEC 61131-3. *)
FUNCTION_BLOCK Shape
  VAR_OUTPUT calls : INT; END_VAR
  METHOD Area : REAL
    Area := 0.0;
  END_METHOD
  METHOD Describe : INT
    Describe := THIS^.Kind();
  END_METHOD
  METHOD Kind : INT
    Kind := 1;
  END_METHOD
  METHOD Twice : INT
    Twice := Kind() * 2;
  END_METHOD
  calls := calls + 1;
END_FUNCTION_BLOCK

FUNCTION_BLOCK Square EXTENDS Shape
  VAR_INPUT side : REAL; END_VAR
  METHOD Area : REAL
    Area := side * side + SUPER^.Area();
  END_METHOD
  METHOD Kind : INT
    Kind := 2;
  END_METHOD
  SUPER^();
END_FUNCTION_BLOCK

PROGRAM main
  VAR sq : Square; END_VAR
  VAR a AT %QD0 : REAL; k AT %QW4 : INT; c AT %QW6 : INT; t AT %QW8 : INT; END_VAR
  sq(side := 3.0);
  a := sq.Area();
  k := sq.Describe();
  c := sq.calls;
  t := sq.Twice();
END_PROGRAM

CONFIGURATION cf
  RESOURCE r ON x
    TASK tk(INTERVAL := T#10ms, PRIORITY := 1);
    PROGRAM p WITH tk : main;
  END_RESOURCE
END_CONFIGURATION

(* ---- codesyspointernumber.st ---- *)
(* A pointer converted to a ULINT or LWORD (pointers, W0017): a number
   naming the place it points at, 0 for NULL - as TcOpen's TcoObject
   keeps `_Identity := ADR(THIS^)` and compares identities. The numbers
   are addresses, so only how they compare is traced:
   ADR(x) twice, once through p: equal (%QX0.0).
   ADR(x) and ADR(y): not equal (%QX0.1).
   NULL: 0 (%QX0.2).
   ADR(THIS^) in a's method, and ADR(a) outside: equal (%QX0.3).
   a's and b's: not equal (%QX0.4).
   As an LWORD, the same number as the ULINT (%QX0.5).
   reference-skip: not IEC 61131-3. *)
FUNCTION_BLOCK Obj
  VAR id : ULINT; END_VAR
  METHOD Identity : ULINT
    id := ADR(THIS^);
    Identity := id;
  END_METHOD
END_FUNCTION_BLOCK

PROGRAM main
  VAR
    x : INT; y : INT; p : POINTER TO INT; n : POINTER TO INT;
    i1 : ULINT; i2 : ULINT; i3 : ULINT; z : ULINT; w : LWORD;
    a : Obj; b : Obj;
  END_VAR
  VAR
    q0 AT %QX0.0 : BOOL; q1 AT %QX0.1 : BOOL; q2 AT %QX0.2 : BOOL;
    q3 AT %QX0.3 : BOOL; q4 AT %QX0.4 : BOOL; q5 AT %QX0.5 : BOOL;
  END_VAR
  p := ADR(x);
  i1 := ADR(x);
  i2 := p;
  i3 := ADR(y);
  z := n;
  w := p;
  q0 := i1 = i2;
  q1 := i1 <> i3;
  q2 := z = 0;
  i1 := ADR(a);
  q3 := a.Identity() = i1;
  q4 := a.Identity() <> b.Identity();
  q5 := LWORD_TO_ULINT(w) = i2;
END_PROGRAM

CONFIGURATION cf
  RESOURCE r ON x
    TASK tk(INTERVAL := T#10ms, PRIORITY := 1);
    PROGRAM p WITH tk : main;
  END_RESOURCE
END_CONFIGURATION

(* ---- codesysprop.st ---- *)
(* CODESYS's PROPERTY (properties), as TcOpen writes them. Worked by hand:
   %QW0: m.Speed := 150, the SET clamps it to 100; read back: 100.
   %QW2: m.Speed := 40, then Boost, inside Motor, Speed := Speed + 5
   through the property itself: 45.
   %QW4: Sets, read only, counts the SET's three calls: 3.
   %QW6: Level through the interface IHasLevel, Speed / 10: 4.
   %QW8: a STRING property: Name := 'xy', its GET adds '!', Twice reads
   THIS^.Name: LEN('xy!') * 2 = 6 (with codesys-oo).
   %QW10, %QW12: Status, a REFERENCE TO a structure (with reference-to),
   written through: Run twice adds 1 to state, 2; d.Status.n := 7, 7.
   %QW14: Limit, a REFERENCE TO INT with no SET, assigned whole through
   its GET: d.Limit := 12, then Bump, inside Dev, Limit := Limit + 30:
   42.
   reference-skip: not IEC 61131-3. *)
INTERFACE IHasLevel
  PROPERTY Level : INT
    GET
    END_GET
  END_PROPERTY
END_INTERFACE

FUNCTION_BLOCK Motor IMPLEMENTS IHasLevel
  VAR _speed : INT; _sets : INT; END_VAR
  PROPERTY PUBLIC Speed : INT
    GET
      Speed := _speed;
    END_GET
    SET
      _sets := _sets + 1;
      IF Speed > 100 THEN
        _speed := 100;
      ELSE
        _speed := Speed;
      END_IF;
    END_SET
  END_PROPERTY
  PROPERTY PUBLIC Sets : INT
    GET
      Sets := _sets;
    END_GET
  END_PROPERTY
  PROPERTY PUBLIC Level : INT
    GET
      Level := Speed / 10;
    END_GET
  END_PROPERTY
  METHOD PUBLIC Boost
    Speed := Speed + 5;
  END_METHOD
END_FUNCTION_BLOCK

FUNCTION_BLOCK Named
  VAR _n : STRING := 'abc'; END_VAR
  PROPERTY PUBLIC Name : STRING
    GET
      Name := CONCAT(_n, '!');
    END_GET
    SET
      _n := Name;
    END_SET
  END_PROPERTY
  METHOD PUBLIC Twice : INT
    Twice := LEN(THIS^.Name) * 2;
  END_METHOD
END_FUNCTION_BLOCK

TYPE St : STRUCT state : INT; n : INT; END_STRUCT; END_TYPE

FUNCTION_BLOCK Dev
  VAR _st : St; _limit : INT; END_VAR
  PROPERTY PUBLIC Limit : REFERENCE TO INT
    GET
      Limit REF= _limit;
    END_GET
  END_PROPERTY
  METHOD PUBLIC Bump
    Limit := Limit + 30;
  END_METHOD
  PROPERTY PUBLIC Status : REFERENCE TO St
    GET
      Status REF= _st;
    END_GET
  END_PROPERTY
  METHOD PUBLIC Run
    Status.state := Status.state + 1;
  END_METHOD
END_FUNCTION_BLOCK

PROGRAM main
  VAR m : Motor; i : IHasLevel; nm : Named; d : Dev; END_VAR
  VAR q0 AT %QW0 : INT; q1 AT %QW2 : INT; q2 AT %QW4 : INT; q3 AT %QW6 : INT; q4 AT %QW8 : INT; q5 AT %QW10 : INT; q6 AT %QW12 : INT; q7 AT %QW14 : INT; END_VAR
  m.Speed := 150;
  q0 := m.Speed;
  m.Speed := 40;
  m.Boost();
  q1 := m.Speed;
  q2 := m.Sets;
  i := m;
  q3 := i.Level;
  nm.Name := 'xy';
  q4 := nm.Twice();
  d.Run();
  d.Run();
  d.Status.n := 7;
  q5 := d.Status.state;
  q6 := d.Status.n;
  d.Limit := 12;
  d.Bump();
  q7 := d.Limit;
END_PROGRAM

CONFIGURATION cf
  RESOURCE r ON x
    TASK tk(INTERVAL := T#10ms, PRIORITY := 1);
    PROGRAM p WITH tk : main;
  END_RESOURCE
END_CONFIGURATION

(* ---- codesysptrcompare.st ---- *)
(* pointers: a pointer given as an input kept in a VAR only assigned and
   compared with <> (W0018), as TcOpen's TcoSignalInfo remembers which
   signal it last looked up.
   Worked by hand, n counting the changes: tick 0: Get(ADR(g)) n 1,
   Get(ADR(g)) the same, n 1; Get(ADR(h)) n 2. Tick 1: Get(ADR(h)) the
   same, n 2; Get(ADR(g)) n 3; Get(ADR(g)) n 3.
   %QW0 2, then 3.
   reference-skip: not IEC 61131-3. *)
FUNCTION_BLOCK Info
  VAR pLast : POINTER TO INT; END_VAR
  VAR_OUTPUT n : INT; END_VAR
  METHOD PUBLIC Get
    VAR_INPUT p : POINTER TO INT; END_VAR
    IF pLast <> p THEN
      n := n + 1;
      pLast := p;
    END_IF;
  END_METHOD
END_FUNCTION_BLOCK

PROGRAM main
  VAR i : Info; g : INT; h : INT; t : INT; END_VAR
  VAR q0 AT %QW0 : INT; END_VAR
  IF t = 0 THEN
    i.Get(p := ADR(g));
    i.Get(p := ADR(g));
    i.Get(p := ADR(h));
  ELSE
    i.Get(p := ADR(h));
    i.Get(p := ADR(g));
    i.Get(p := ADR(g));
  END_IF;
  t := t + 1;
  q0 := i.n;
END_PROGRAM

CONFIGURATION cf
  RESOURCE r ON x
    TASK tk(INTERVAL := T#10ms, PRIORITY := 1);
    PROGRAM p WITH tk : main;
  END_RESOURCE
END_CONFIGURATION

(* ---- codesysqueryitf.st ---- *)
(* CODESYS's __QUERYINTERFACE (query-interface), as TcOpen asks its
   parent for a drive: `__QUERYINTERFACE(Parent, d)` is `d ?= Parent`,
   TRUE when d then holds the instance. Worked by hand:
   %QW0 the motor implements IDrive: TRUE, its Speed 7: 7.
   %QW2 the lamp does not: FALSE, -1; and d, which held the motor, is
        NULL after: + 100, 99.
   %QW4 no parent: FALSE, 0 stays.
   %QW6 a lamp's derived type implements IDrive, asked through IObj:
        its Speed 42.
   %QW8 in an expression, ANDed with what reads d after it: TRUE AND
        TRUE, 10; the lamp's FALSE, and d NULL after it, 1: 11.
   reference-skip: not IEC 61131-3. *)
INTERFACE IObj EXTENDS __SYSTEM.IQueryInterface
  METHOD Id : INT
  END_METHOD
END_INTERFACE

INTERFACE IDrive EXTENDS __System.IQueryInterface
  METHOD Speed : INT
  END_METHOD
END_INTERFACE

FUNCTION_BLOCK Motor IMPLEMENTS IObj, IDrive
  METHOD PUBLIC Id : INT
    Id := 1;
  END_METHOD
  METHOD PUBLIC Speed : INT
    Speed := 7;
  END_METHOD
END_FUNCTION_BLOCK

FUNCTION_BLOCK Lamp IMPLEMENTS IObj
  METHOD PUBLIC Id : INT
    Id := 2;
  END_METHOD
END_FUNCTION_BLOCK

FUNCTION_BLOCK FastLamp EXTENDS Lamp IMPLEMENTS IDrive
  METHOD PUBLIC Speed : INT
    Speed := 42;
  END_METHOD
END_FUNCTION_BLOCK

FUNCTION_BLOCK Child
  VAR_INPUT Parent : IObj; END_VAR
  VAR_OUTPUT q : INT; END_VAR
  VAR d : IDrive; END_VAR
  IF __QUERYINTERFACE(THIS^.Parent, d) THEN
    q := d.Speed();
  ELSE
    q := -1;
  END_IF
END_FUNCTION_BLOCK

PROGRAM main
  VAR m : Motor; l : Lamp; f : FastLamp; c : Child; o : IObj; d : IDrive; ok : BOOL; END_VAR
  VAR q0 AT %QW0 : INT; q2 AT %QW2 : INT; q4 AT %QW4 : INT; q6 AT %QW6 : INT; q8 AT %QW8 : INT; END_VAR
  c(Parent := m);
  q0 := c.q;
  o := l;
  d := m;
  IF __QUERYINTERFACE(o, d) THEN
    q2 := 1;
  ELSE
    q2 := -1;
  END_IF
  IF d = NULL THEN
    q2 := q2 + 100;
  END_IF
  o := NULL;
  IF __QUERYINTERFACE(o, d) THEN
    q4 := 1;
  END_IF
  c(Parent := f);
  q6 := c.q;
  o := m;
  ok := __QUERYINTERFACE(o, d) AND d.Speed() = 7;
  q8 := 10 * BOOL_TO_INT(ok);
  o := l;
  ok := NOT __QUERYINTERFACE(o, d) AND d = NULL;
  q8 := q8 + BOOL_TO_INT(ok);
END_PROGRAM

CONFIGURATION cf
  RESOURCE r ON x
    TASK tk(INTERVAL := T#10ms, PRIORITY := 1);
    PROGRAM p WITH tk : main;
  END_RESOURCE
END_CONFIGURATION

(* ---- codesysreads.st ---- *)
(* A function block's internal VAR read from outside, never written
   (internal-reads), as CODESYS and TwinCAT allow, each read warned
   (W0012). Worked by hand, after a(x := 5) and a(x := 6):
   %QW0: a.count, 2.  %QD2: a.total, 5 + 6 = 11.
   %QW6: a.arr[2], 3.  %QW8: a.inn.q, Inner's output, 7.
   %QW10: a.inn.k, Inner's own VAR, 7.
   %QW12: dr.st.Restore() twice, a method of Drive's internal instance
   st, as TcOpen calls one: 10 + 10 = 20.
   %QW14: dr.cnt(inc := 3, total => q6) twice, Drive's internal
   instance cnt called from outside, as TcOpen's `_failTimer(...)`
   through its task: 3 + 3 = 6. %QW16: w.dr.cnt(inc := 100) once,
   two levels in, then w.dr.cnt.total read: 100.
   reference-skip: not IEC 61131-3. *)
FUNCTION_BLOCK Inner
  VAR_OUTPUT q : INT; END_VAR
  VAR k : INT := 7; END_VAR
  q := k;
END_FUNCTION_BLOCK

FUNCTION_BLOCK Acc
  VAR_INPUT x : INT; END_VAR
  VAR count : INT; total : DINT; arr : ARRAY[0..2] OF INT := [1, 2, 3]; inn : Inner; END_VAR
  count := count + 1;
  total := total + x;
  inn();
END_FUNCTION_BLOCK

FUNCTION_BLOCK State
  VAR_OUTPUT n : INT; END_VAR
  METHOD PUBLIC Restore
    n := n + 10;
  END_METHOD
END_FUNCTION_BLOCK

FUNCTION_BLOCK Counter
  VAR_INPUT inc : INT; END_VAR
  VAR_OUTPUT total : INT; END_VAR
  total := total + inc;
END_FUNCTION_BLOCK

FUNCTION_BLOCK Drive
  VAR st : State; cnt : Counter; END_VAR
END_FUNCTION_BLOCK

FUNCTION_BLOCK Wrap
  VAR dr : Drive; END_VAR
END_FUNCTION_BLOCK

PROGRAM main
  VAR a : Acc; dr : Drive; w : Wrap; END_VAR
  VAR q0 AT %QW0 : INT; q1 AT %QD2 : DINT; q2 AT %QW6 : INT; q3 AT %QW8 : INT; q4 AT %QW10 : INT; q5 AT %QW12 : INT;
      q6 AT %QW14 : INT; q7 AT %QW16 : INT; END_VAR
  a(x := 5);
  a(x := 6);
  q0 := a.count;
  q1 := a.total;
  q2 := a.arr[2];
  q3 := a.inn.q;
  q4 := a.inn.k;
  dr.st.Restore();
  dr.st.Restore();
  q5 := dr.st.n;
  dr.cnt(inc := 3, total => q6);
  dr.cnt(inc := 3, total => q6);
  w.dr.cnt(inc := 100);
  q7 := w.dr.cnt.total;
END_PROGRAM

CONFIGURATION cf
  RESOURCE r ON x
    TASK tk(INTERVAL := T#10ms, PRIORITY := 1);
    PROGRAM p WITH tk : main;
  END_RESOURCE
END_CONFIGURATION

(* ---- codesysrefthis.st ---- *)
(* A method that gives its own instance as a REFERENCE TO, `REF= THIS^`,
   called again on what it gives - TcOpen's StringBuilder,
   `sb.Append('a').Append('b')` (codesys-oo, reference-to).
   twice overrides add: a call through the reference given reaches it.
   Worked by hand, each tick:
   a.add(1).add(2).add(3): a.n + 6.
   t.add(1).add(10): twice's both, + 2 + 20; r REF= t.add(100): + 200,
   r is t; r.add(1000), through r, twice's: + 2000. t.n + 2222.
   %QD0 a.n, %QD4 t.n, %QD8 r.n (t's):
   tick 0: 6, 2222, 2222; tick 1: 12, 4444, 4444.
   reference-skip: not IEC 61131-3. *)
FUNCTION_BLOCK acc
  VAR_OUTPUT n : DINT; END_VAR
  METHOD add : REFERENCE TO acc
    VAR_INPUT k : DINT; END_VAR
    n := n + k;
    add REF= THIS^;
  END_METHOD
END_FUNCTION_BLOCK

FUNCTION_BLOCK twice EXTENDS acc
  METHOD add : REFERENCE TO acc
    VAR_INPUT k : DINT; END_VAR
    n := n + 2 * k;
    add REF= THIS^;
  END_METHOD
END_FUNCTION_BLOCK

PROGRAM main
  VAR a : acc; t : twice; r : REFERENCE TO acc; END_VAR
  VAR q0 AT %QD0 : DINT; END_VAR
  VAR q1 AT %QD4 : DINT; END_VAR
  VAR q2 AT %QD8 : DINT; END_VAR
  a.add(1).add(2).add(3);
  t.add(1).add(10);
  r REF= t.add(100);
  r.add(1000);
  q0 := a.n;
  q1 := t.n;
  q2 := r.n;
END_PROGRAM

CONFIGURATION cf
  RESOURCE r ON x
    TASK tk(INTERVAL := T#10ms, PRIORITY := 1);
    PROGRAM p WITH tk : main;
  END_RESOURCE
END_CONFIGURATION

(* ---- codesysshortcircuit.st ---- *)
(* AND_THEN and OR_ELSE (short-circuit): the right operand evaluated
   only when the left does not decide, as CODESYS and TwinCAT have them.
   c.Hit() counts its calls. Worked by hand:
   cycle 0: FALSE AND_THEN c.Hit(): not called, FALSE; TRUE AND_THEN
     c.Hit(): called (n 1), TRUE; TRUE OR_ELSE c.Hit(): not called, TRUE;
     FALSE OR_ELSE c.Hit(): called (n 2), TRUE. %QW0 n = 2;
     %QW2 r1 + 2 r2 + 4 r3 + 8 r4 = 0 + 2 + 4 + 8 = 14.
     d = 0: d <> 0 AND_THEN 10 / d > 1 divides not, no fault: %QW4 7.
     The same in an IF's ELSIF and a WHILE, each Hit() a call more only
     where the left lets it: k 1 (ELSIF taken), %QW6 = n after = 3.
   cycle 1: n from 3: 5, 14, 7; %QW6 6.
   reference-skip: not IEC 61131-3. *)
FUNCTION_BLOCK Counter
VAR_OUTPUT n : INT; END_VAR
METHOD PUBLIC Hit : BOOL
n := n + 1;
Hit := TRUE;
END_METHOD
END_FUNCTION_BLOCK

PROGRAM main
  VAR c : Counter; f : BOOL; t : BOOL := TRUE; r1, r2, r3, r4 : BOOL; d, k : INT; END_VAR
  VAR q AT %QW0 : INT; x AT %QW2 : INT; w AT %QW4 : INT; v AT %QW6 : INT; END_VAR
  r1 := f AND_THEN c.Hit();
  r2 := t AND_THEN c.Hit();
  r3 := t OR_ELSE c.Hit();
  r4 := f OR_ELSE c.Hit();
  q := c.n;
  x := BOOL_TO_INT(r1) + 2 * BOOL_TO_INT(r2) + 4 * BOOL_TO_INT(r3) + 8 * BOOL_TO_INT(r4);
  w := 0;
  IF d <> 0 AND_THEN 10 / d > 1 THEN
    w := 1;
  END_IF;
  w := w + 7;
  k := 0;
  IF f AND_THEN c.Hit() THEN
    k := 2;
  ELSIF t AND_THEN c.Hit() THEN
    k := 1;
  END_IF;
  WHILE k > 0 AND_THEN t DO
    k := k - 1;
  END_WHILE;
  v := c.n;
END_PROGRAM

CONFIGURATION cf
  RESOURCE r ON x
    TASK tk(INTERVAL := T#10ms, PRIORITY := 1);
    PROGRAM p WITH tk : main;
  END_RESOURCE
END_CONFIGURATION

(* ---- codesysstructblocks.st ---- *)
(* CODESYS's and TwinCAT's structures holding blocks set up by their
   FB_init (struct-blocks), as TcOpen's TcoStruct: an ABSTRACT base
   structure whose member Self is given the structure itself (THIS^),
   a structure extending it whose members are given Self, a sibling.
   Worked by hand, h's d set up with Parent := THIS^ (h) and tag := 5,
   then each member's FB_init in the order declared:
   Self.FB_init(s := d): Self references d.
   a.FB_init(p := Self, k := 1): up := Self.Id(), d.tag + 100 = 105.
   b.FB_init(p := Self, k := 2): n := 2.
   %QW0 d.a.up 105, %QW2 d.b.n 2, %QW4 Self.ParentId(), d.Parent.Id(),
   h's 42, %QW6 Self.Id() 105.
   d.inner, an Inner (a Base too) given Parent := Self, d's own member,
   and tag 9: its c.FB_init(p := inner.Self): 9 + 100, %QW8 109; its
   Self.ParentId() is its Parent's Id, d.Self's, %QW10 105.
   reference-skip: not IEC 61131-3. *)
INTERFACE IObj
  METHOD Id : INT
  END_METHOD
END_INTERFACE

TYPE
  ABSTRACT Base : STRUCT
    Parent : IObj;
    Self : Marker(THIS^);
    tag : INT := 7;
  END_STRUCT;
END_TYPE

TYPE Inner EXTENDS Base :
STRUCT
  c : Leaf(Self, 3);
END_STRUCT
END_TYPE

TYPE Data EXTENDS Base :
STRUCT
  a : Leaf(Self, 1);
  b : Leaf(Self, 2);
  inner : Inner := (Parent := Self, tag := 9);
END_STRUCT
END_TYPE

FUNCTION_BLOCK Marker IMPLEMENTS IObj
  VAR st : REFERENCE TO Base; END_VAR
  METHOD FB_init : BOOL
    VAR_INPUT bInitRetains : BOOL; bInCopyCode : BOOL; s : REFERENCE TO Base; END_VAR
    st REF= s;
  END_METHOD
  METHOD PUBLIC Id : INT
    Id := st.tag + 100;
  END_METHOD
  METHOD PUBLIC ParentId : INT
    ParentId := st.Parent.Id();
  END_METHOD
END_FUNCTION_BLOCK

FUNCTION_BLOCK Leaf
  VAR_OUTPUT up : INT; n : INT; END_VAR
  METHOD FB_init : BOOL
    VAR_INPUT bInitRetains : BOOL; bInCopyCode : BOOL; p : IObj; k : INT; END_VAR
    up := p.Id();
    n := k;
  END_METHOD
END_FUNCTION_BLOCK

FUNCTION_BLOCK Holder IMPLEMENTS IObj
  VAR d : Data := (Parent := THIS^, tag := 5); END_VAR
  VAR_OUTPUT o1 : INT; o2 : INT; o3 : INT; o4 : INT; o5 : INT; o6 : INT; END_VAR
  METHOD PUBLIC Id : INT
    Id := 42;
  END_METHOD
  o1 := d.a.up;
  o2 := d.b.n;
  o3 := d.Self.ParentId();
  o4 := d.Self.Id();
  o5 := d.inner.c.up;
  o6 := d.inner.Self.ParentId();
END_FUNCTION_BLOCK

PROGRAM main
  VAR h : Holder; END_VAR
  VAR q0 AT %QW0 : INT; q1 AT %QW2 : INT; q2 AT %QW4 : INT; q3 AT %QW6 : INT; q4 AT %QW8 : INT;
      q5 AT %QW10 : INT; END_VAR
  h();
  q0 := h.o1; q1 := h.o2; q2 := h.o3; q3 := h.o4; q4 := h.o5; q5 := h.o6;
END_PROGRAM

CONFIGURATION cf
  RESOURCE r ON x
    TASK tk(INTERVAL := T#10ms, PRIORITY := 1);
    PROGRAM p WITH tk : main;
  END_RESOURCE
END_CONFIGURATION

(* ---- codesysstructinout.st ---- *)
(* A structure extending another given to an in-out of its base's type
   (struct-extends), as TcOpen's TcoTixonFeeding gives its steps' Config,
   Control and Status to its tasks' generic in-outs. The block keeps the
   in-out and a method writes through it later (method-in-outs).
   Worked by hand, each tick: bp(io := t) adds 10 to t.a, bp.Again()
   100; F(m := t) adds 5 to t.b and gives t.a + t.b; bq(io := arr[i])
   adds 10 to arr[2].a. Tick 1: t.a 1 + 110 = 111, t.b 2 + 5 = 7,
   F 118, t.c 3, arr[2].a 11, arr[1].a 1. Tick 2: t.a 221, t.b 12,
   F 233, t.c 3, arr[2].a 21, arr[1].a 1.
   reference-skip: not IEC 61131-3. *)
TYPE
  Base : STRUCT a : INT := 1; END_STRUCT;
  Middle EXTENDS Base : STRUCT b : INT := 2; END_STRUCT;
  Top EXTENDS Middle : STRUCT c : INT := 3; END_STRUCT;
END_TYPE

FUNCTION_BLOCK Bump
  VAR_IN_OUT io : Base; END_VAR
  METHOD Again
    io.a := io.a + 100;
  END_METHOD
  io.a := io.a + 10;
END_FUNCTION_BLOCK

FUNCTION F : INT
  VAR_IN_OUT m : Middle; END_VAR
  m.b := m.b + 5;
  F := m.a + m.b;
END_FUNCTION

PROGRAM main
  VAR t : Top; arr : ARRAY[1..2] OF Top; i : INT := 2; bp : Bump; bq : Bump; x : INT; END_VAR
  VAR q0 AT %QW0 : INT; q2 AT %QW2 : INT; q4 AT %QW4 : INT; END_VAR
  VAR q6 AT %QW6 : INT; q8 AT %QW8 : INT; q10 AT %QW10 : INT; END_VAR
  bp(io := t);
  bp.Again();
  x := F(m := t);
  bq(io := arr[i]);
  q0 := t.a;
  q2 := t.b;
  q4 := x;
  q6 := t.c;
  q8 := arr[2].a;
  q10 := arr[1].a;
END_PROGRAM

CONFIGURATION cf
  RESOURCE r ON x
    TASK tk(INTERVAL := T#10ms, PRIORITY := 1);
    PROGRAM p WITH tk : main;
  END_RESOURCE
END_CONFIGURATION

(* ---- codesyssuper.st ---- *)
(* CODESYS's and TwinCAT's SUPER^ (super-calls), as TcOpen writes it.
   Worked by hand, d called once with x = 100:
   SUPER^(i := 3, io := io, o => got): the base's body with i = 3,
   io bound to itself: n 1, o 30, x 103; got 30.
   SUPER^(i := 4), a second call in the body: n 2, o 40, x 107.
   THIS^.Again(), a method calling SUPER^() on i = 4: n 3, o 40, x 111.
   SUPER^.Kind, the base's GET, not Derived's: 1; THIS^.Kind: 2.
   k := SUPER^.n, the instance's own n: 3; SUPER^.n := 10, m := n: 10.
   %QW0 got 30, %QW2 o 40, %QW4 x 111, %QW6 1, %QW8 2, %QW10 3, %QW12 10.
   reference-skip: not IEC 61131-3. *)
FUNCTION_BLOCK Base
  VAR_INPUT i : INT; END_VAR
  VAR_IN_OUT io : INT; END_VAR
  VAR_OUTPUT o : INT; END_VAR
  VAR n : INT; END_VAR
  PROPERTY PUBLIC Kind : INT
    GET
      Kind := 1;
    END_GET
  END_PROPERTY
  n := n + 1;
  o := i * 10;
  io := io + i;
END_FUNCTION_BLOCK

FUNCTION_BLOCK Derived EXTENDS Base
  VAR_OUTPUT got : INT; viaSuper : INT; own : INT; k : INT; m : INT; END_VAR
  PROPERTY PUBLIC Kind : INT
    GET
      Kind := 2;
    END_GET
  END_PROPERTY
  METHOD PUBLIC Again
    SUPER^();
  END_METHOD
  SUPER^(i := 3, io := io, o => got);
  SUPER^(i := 4);
  THIS^.Again();
  viaSuper := SUPER^.Kind;
  own := THIS^.Kind;
  k := SUPER^.n;
  SUPER^.n := 10;
  m := n;
END_FUNCTION_BLOCK

PROGRAM main
  VAR d : Derived; x : INT := 100; END_VAR
  VAR
    q0 AT %QW0 : INT; q1 AT %QW2 : INT; q2 AT %QW4 : INT; q3 AT %QW6 : INT;
    q4 AT %QW8 : INT; q5 AT %QW10 : INT; q6 AT %QW12 : INT;
  END_VAR
  d(io := x);
  q0 := d.got; q1 := d.o; q2 := x; q3 := d.viaSuper; q4 := d.own; q5 := d.k; q6 := d.m;
END_PROGRAM

CONFIGURATION cf
  RESOURCE r ON x
    TASK tk(INTERVAL := T#10ms, PRIORITY := 1);
    PROGRAM p WITH tk : main;
  END_RESOURCE
END_CONFIGURATION

(* ---- codesysthisinit.st ---- *)
(* CODESYS's and TwinCAT's THIS^ in an initial value (codesys-oo), as
   TcOpen writes `(Parent := THIS^)`: each instance's structure holds
   that instance, through the interface. Worked by hand:
   %QW0 a.Ask(): a's Id, k 1, plus n 5: 6.
   %QW2 b.Ask(): b's own Parent, not a's: 2 + 5, 7.
   %QW4 s.Ask(): s is a Special, whose Id overrides: 3 * 100 + 5, 305.
   reference-skip: not IEC 61131-3. *)
INTERFACE IObj
  METHOD Id : INT
  END_METHOD
END_INTERFACE

TYPE
  Holder : STRUCT
    Parent : IObj;
    n : INT;
  END_STRUCT;
END_TYPE

FUNCTION_BLOCK Comp IMPLEMENTS IObj
  VAR_INPUT k : INT; END_VAR
  VAR h : Holder := (Parent := THIS^, n := 5); END_VAR
  METHOD PUBLIC Id : INT
    Id := k;
  END_METHOD
  METHOD PUBLIC Ask : INT
    Ask := h.Parent.Id() + h.n;
  END_METHOD
END_FUNCTION_BLOCK

FUNCTION_BLOCK Special EXTENDS Comp
  METHOD PUBLIC Id : INT
    Id := k * 100;
  END_METHOD
END_FUNCTION_BLOCK

PROGRAM main
  VAR a : Comp; b : Comp; s : Special; END_VAR
  VAR qa AT %QW0 : INT; qb AT %QW2 : INT; qs AT %QW4 : INT; END_VAR
  a(k := 1);
  b(k := 2);
  s(k := 3);
  qa := a.Ask();
  qb := b.Ask();
  qs := s.Ask();
END_PROGRAM

CONFIGURATION cf
  RESOURCE r ON x
    TASK tk(INTERVAL := T#10ms, PRIORITY := 1);
    PROGRAM p WITH tk : main;
  END_RESOURCE
END_CONFIGURATION

(* ---- codesystypeconst.st ---- *)
(* A block's constant read through its type's name (type-constants), as
   TcOpen sizes its messages' strings by TcoMessengerEnv's. Worked by
   hand: Env.N 8, Env.TWICE N * 2 = 16.
   %QW0 Env.TWICE + the upper bound of a, ARRAY[1..Env.TWICE]: 32;
   %QW2 s, a STRING[Env.N], given 11 characters: cut to 8 (flagged), LEN 8;
   %QW4 Env.HALF, an LREAL 3.5, * 2: 7. The same each cycle.
   reference-skip: not IEC 61131-3. *)
FUNCTION_BLOCK Env
VAR CONSTANT
  N : INT := 8;
  TWICE : INT := N * 2;
  HALF : LREAL := 3.5;
END_VAR
END_FUNCTION_BLOCK

PROGRAM main
  VAR s : STRING[Env.N]; a : ARRAY[1..Env.TWICE] OF INT; END_VAR
  VAR x AT %QW0 : INT; y AT %QW2 : INT; z AT %QW4 : INT; END_VAR
  x := Env.TWICE + DINT_TO_INT(UPPER_BOUND(a, 1));
  s := 'abcdefghijk';
  y := LEN(s);
  z := LREAL_TO_INT(Env.HALF * 2.0);
END_PROGRAM

CONFIGURATION cf
  RESOURCE r ON x
    TASK tk(INTERVAL := T#10ms, PRIORITY := 1);
    PROGRAM p WITH tk : main;
  END_RESOURCE
END_CONFIGURATION

(* ---- codesysvarinfo.st ---- *)
(* CODESYS's and TwinCAT's __VARINFO (var-info): a __SYSTEM.VAR_INFO of
   a variable, as TcOpen's tasks name the signal they wait for in a
   message (`__VARINFO(inoStatus.State...).Symbol`).
   Worked by hand, the same each tick:
   %QB0 LEN(msg), 'waiting for ' (12) + 'ES_IsStopped' (12): 24;
   %QB1 BitSize of a BOOL, a byte: 8;
   %QB2 TypeClass of io.Vals is TYPE_ARRAY: 1;
   %QB3 NumElements of ARRAY[1..3] OF INT: 3;
   %QB4 ElemBitSize, an INT: 16;
   %QB5 BaseTypeClass is TYPE_INT: 1;
   %QB6 LEN(TypeName), 'ARRAY[1..3] OF INT': 18;
   %QB7 BitNo of w.5: 5; %QB8 its BitSize: 1;
   %QB9 MemoryArea, CODESYS's initial MEM_MEMORY: 1.
   reference-skip: not IEC 61131-3. *)
TYPE Sig : STRUCT
  ES_IsStopped : BOOL;
  Vals : ARRAY[1..3] OF INT;
END_STRUCT;
END_TYPE

FUNCTION_BLOCK Watch
  VAR_IN_OUT io : Sig; END_VAR
  VAR_OUTPUT msg : STRING[60]; bits : INT; END_VAR
  VAR info : __SYSTEM.VAR_INFO; END_VAR
  info := __VARINFO(io.ES_IsStopped);
  msg := CONCAT('waiting for ', info.Symbol);
  bits := info.BitSize;
END_FUNCTION_BLOCK

PROGRAM main
  VAR s : Sig; wt : Watch; info : __SYSTEM.VAR_INFO; w : WORD; END_VAR
  VAR q AT %QB0 : ARRAY[0..9] OF BYTE; END_VAR
  wt(io := s);
  q[0] := TO_BYTE(LEN(wt.msg));
  q[1] := TO_BYTE(wt.bits);
  info := __VARINFO(s.Vals);
  q[2] := BOOL_TO_BYTE(info.TypeClass = __SYSTEM.TYPE_CLASS.TYPE_ARRAY);
  q[3] := TO_BYTE(info.NumElements);
  q[4] := TO_BYTE(info.ElemBitSize);
  q[5] := BOOL_TO_BYTE(info.BaseTypeClass = __SYSTEM.TYPE_CLASS.TYPE_INT);
  q[6] := TO_BYTE(LEN(info.TypeName));
  info := __VARINFO(w.5);
  q[7] := TO_BYTE(info.BitNo);
  q[8] := TO_BYTE(info.BitSize);
  q[9] := BOOL_TO_BYTE(info.MemoryArea = __SYSTEM.MEMORY_AREA.MEM_MEMORY);
END_PROGRAM

CONFIGURATION cf
  RESOURCE r ON x
    TASK tk(INTERVAL := T#10ms, PRIORITY := 1);
    PROGRAM p WITH tk : main;
  END_RESOURCE
END_CONFIGURATION

(* ---- codesysvarinst.st ---- *)
(* A method's instance variables (var-inst), as TcOpen's messenger keeps
   the cycle its StringBuilder was last read in: one for each instance,
   set up once, kept from call to call. Worked by hand, two instances:
   cycle 0: a.Next() 10 -> 11, a.Next() 12; b.Next() 11: own count;
     a.Calls (a property's GET counting its reads) 1, b.Calls 1:
     %QW0 a.Next 12, %QW2 b 11, %QW4 a.Calls + 10 * b.Calls 11;
     d, derived, its own from 10: %QW6 11.
   cycle 1: a 13, 14; b 12; Calls 2 and 2: 22; d 12.
   reference-skip: not IEC 61131-3. *)
FUNCTION_BLOCK Seq
METHOD PUBLIC Next : INT
VAR_INST
  n : INT := 10;
END_VAR
n := n + 1;
Next := n;
END_METHOD
PROPERTY PUBLIC Calls : INT
GET
VAR_INST
  reads : INT;
END_VAR
reads := reads + 1;
Calls := reads;
END_GET
END_PROPERTY
END_FUNCTION_BLOCK

FUNCTION_BLOCK Derived EXTENDS Seq
END_FUNCTION_BLOCK

PROGRAM main
  VAR a, b : Seq; d : Derived; t : INT; END_VAR
  VAR x AT %QW0 : INT; y AT %QW2 : INT; z AT %QW4 : INT; w AT %QW6 : INT; END_VAR
  t := a.Next();
  x := a.Next();
  y := b.Next();
  z := a.Calls + 10 * b.Calls;
  w := d.Next();
END_PROGRAM

CONFIGURATION cf
  RESOURCE r ON x
    TASK tk(INTERVAL := T#10ms, PRIORITY := 1);
    PROGRAM p WITH tk : main;
  END_RESOURCE
END_CONFIGURATION

(* ---- codesysvarstat.st ---- *)
(* Static variables (var-stat), as TcOpen's messenger and CRC blocks
   declare them: one of each for the POU, shared by every instance and
   kept from call to call. Worked by hand, two cycles:
   cycle 0: a() n 5 -> 6, b() 7; a.Bump() k 1, n 17; b.Bump() k 2, n 27:
     %QW0 x = 1 + 2 = 3; F twice through its loop: %QW2 2;
     m(), More's body only: %QW4 r = 27 * 2 = 54; %QW6 a.q = 6.
   cycle 1: a() 28, b() 29; Bump 3 (n 39), 4 (n 49): %QW0 7;
     F: %QW2 4; %QW4 98; %QW6 28.
   reference-skip: not IEC 61131-3. *)
FUNCTION_BLOCK Cnt
VAR_STAT
  n : INT := 5;
END_VAR
VAR_OUTPUT q : INT; END_VAR
METHOD PUBLIC Bump : INT
VAR_STAT k : INT; END_VAR
k := k + 1;
n := n + 10;
Bump := k;
END_METHOD
n := n + 1;
q := n;
END_FUNCTION_BLOCK

FUNCTION_BLOCK More EXTENDS Cnt
VAR_OUTPUT r : INT; END_VAR
r := n * 2;
END_FUNCTION_BLOCK

FUNCTION F : INT
VAR_STAT calls : INT; i : INT; END_VAR
FOR i := 1 TO 2 DO
  calls := calls + 1;
END_FOR;
F := calls;
END_FUNCTION

PROGRAM main
  VAR a, b : Cnt; m : More; END_VAR
  VAR x AT %QW0 : INT; y AT %QW2 : INT; z AT %QW4 : INT; w AT %QW6 : INT; END_VAR
  a();
  b();
  x := a.Bump() + b.Bump();
  y := F();
  m();
  z := m.r;
  w := a.q;
END_PROGRAM

CONFIGURATION cf
  RESOURCE r ON x
    TASK tk(INTERVAL := T#10ms, PRIORITY := 1);
    PROGRAM p WITH tk : main;
  END_RESOURCE
END_CONFIGURATION

(* ---- confignest.st ---- *)
(* VAR_CONFIG's initial value for a variable of a block held in a
   RETAIN block (Ed.3 6.5.6.2, 6.8.2): the inner block is in a section
   that says neither RETAIN nor NON_RETAIN, so it keeps what its own
   type says, nothing, and starts again at a warm restart - with
   VAR_CONFIG's value, which prevails. Worked by hand:

   tick 0: b.x 50 + 1 = 51 (Q0 33 00); a.y 70 + 1 = 71 (Q2 47 00).
   tick 1: 52, 72.
   warm, before tick 2: a is RETAIN, y stays 72; b starts again, x 1,
   then VAR_CONFIG's 50.
   tick 2: 51 (33 00), 73 (49 00).
   confignest.iecf.trace: the reference compiler generates nothing for
   VAR_CONFIG (as `varconfig`), and its host's warm restart is a cold
   one: x and y from 1 each time. *)
FUNCTION_BLOCK inner
  VAR_OUTPUT x : INT := 1; END_VAR
  x := x + 1;
END_FUNCTION_BLOCK
FUNCTION_BLOCK outer
  VAR_OUTPUT y : INT := 1; END_VAR
  VAR b : inner; END_VAR
  VAR_OUTPUT bx : INT; END_VAR
  b();
  y := y + 1;
  bx := b.x;
END_FUNCTION_BLOCK
PROGRAM main
  VAR RETAIN a : outer; END_VAR
  VAR q AT %QW0 : INT; q2 AT %QW2 : INT; END_VAR
  a();
  q := a.bx;
  q2 := a.y;
END_PROGRAM
CONFIGURATION plant
  RESOURCE cpu ON PLC
    TASK t(INTERVAL := T#10ms, PRIORITY := 1);
    PROGRAM p WITH t : main;
  END_RESOURCE
  VAR_CONFIG
    cpu.p.a.b.x : INT := 50;
    cpu.p.a.y : INT := 70;
  END_VAR
END_CONFIGURATION

(* ---- connect2.st ---- *)
(* A program's connections (Ed.3 6.8.2) of strings, subranges, fields,
   and in-outs of every kind: a structure, an array, a STRING, an
   instance, variables at addresses, a subrange of other bounds.
   Worked by hand, tick 0 then tick 1:
   s : STRING[3] := 'abcdef' is cut: LEN 3 (%QB0); flagged
   STRING_LENGTH, the first flag, at the CONFIGURATION's line of it.
   a : SUBR (0..5) := 9 is clamped: 5 (%QB1). f := gp.x, a field: 7,
   then 8 (%QB2). o => gsub, a SUBR, given 9: 5, read through gsub the
   next tick: 0 then 5 (%QB3). os => gs2, a STRING[2], given 'abcd':
   'ab', LEN 0 then 2 (%QB4).
   In-outs, the globals themselves: ip.x + 1, gp.x 8 then 9 (%QB5);
   ia[2] + 10, ga[2] 12 then 22 (%QB6); is + 'z', gstr 'az' then 'azz'
   (%QB7); ic(), gcnt.n 1 then 2 (%QB8).
   At addresses, copied in before the run and back after it: il, gl at
   %MW0, 4 + 1 = 5 then 6 (%QB9, and %MW0); ila[1], gla at %MW2, 10 + 2
   = 12 then 14 (%QB10, and %MW2).
   isub, an INT, given gsub2, a SUBR of 1: 1 + 9 = 10 in the program
   (%QB11), stored back clamped to 5; the next tick 5 + 9 = 14.
   reference-skip: the reference compiler crashes on program
   connections (connections). *)
TYPE
  SUBR : INT (0..5);
  PT : STRUCT x : INT; END_STRUCT;
END_TYPE
FUNCTION_BLOCK Cnt
  VAR_OUTPUT n : INT; END_VAR
  n := n + 1;
END_FUNCTION_BLOCK
PROGRAM main
  VAR_INPUT s : STRING[3]; a : SUBR; f : INT; END_VAR
  VAR_OUTPUT o : INT; os : STRING; END_VAR
  VAR_IN_OUT
    ip : PT;
    ia : ARRAY [1..3] OF INT;
    is : STRING;
    ic : Cnt;
    il : INT;
    ila : ARRAY [1..2] OF INT;
    isub : INT;
  END_VAR
  VAR_EXTERNAL gsub : SUBR; gs2 : STRING[2]; END_VAR
  VAR
    q0 AT %QB0 : SINT;
    q1 AT %QB1 : SINT;
    q2 AT %QB2 : SINT;
    q3 AT %QB3 : SINT;
    q4 AT %QB4 : SINT;
    q5 AT %QB5 : SINT;
    q6 AT %QB6 : SINT;
    q7 AT %QB7 : SINT;
    q8 AT %QB8 : SINT;
    q9 AT %QB9 : SINT;
    q10 AT %QB10 : SINT;
    q11 AT %QB11 : SINT;
  END_VAR
  q0 := INT_TO_SINT(LEN(s));
  q1 := INT_TO_SINT(a);
  q2 := INT_TO_SINT(f);
  q3 := INT_TO_SINT(gsub);
  q4 := INT_TO_SINT(LEN(gs2));
  ip.x := ip.x + 1;
  q5 := INT_TO_SINT(ip.x);
  ia[2] := ia[2] + 10;
  q6 := INT_TO_SINT(ia[2]);
  is := CONCAT(is, 'z');
  q7 := INT_TO_SINT(LEN(is));
  ic();
  q8 := INT_TO_SINT(ic.n);
  il := il + 1;
  q9 := INT_TO_SINT(il);
  ila[1] := ila[1] + 2;
  q10 := INT_TO_SINT(ila[1]);
  isub := isub + 9;
  q11 := INT_TO_SINT(isub);
  o := 9;
  os := 'abcd';
END_PROGRAM

CONFIGURATION c
  VAR_GLOBAL
    gp : PT := (x := 7);
    ga : ARRAY [1..3] OF INT := [1, 2, 3];
    gstr : STRING := 'a';
    gcnt : Cnt;
    gsub : SUBR;
    gs2 : STRING[2];
    gsub2 : SUBR := 1;
  END_VAR
  VAR_GLOBAL
    gl AT %MW0 : INT := 4;
    gla AT %MW2 : ARRAY [1..2] OF INT := [10, 20];
  END_VAR
  RESOURCE r ON x
    TASK t(INTERVAL := T#10ms, PRIORITY := 1);
    PROGRAM p WITH t : main(
      s := 'abcdef',
      a := 9,
      f := gp.x,
      o => gsub,
      os => gs2,
      ip := gp,
      ia := ga,
      is := gstr,
      ic := gcnt,
      il := gl,
      ila := gla,
      isub := gsub2);
  END_RESOURCE
END_CONFIGURATION

(* ---- constfns.st ---- *)
(* Initial values that are standard functions of constants (Ed.3
   6.6.1.2.4): worked out by the compiler where the result is exact,
   and the mathematics of Table 28 and ** computed as the variable is
   set up, by the target's own, once the compiler has worked out that
   the result is one the type holds - in a program, a TYPE, a
   structure's field, an array, a global, a block's input and a
   FUNCTION's input and own variable.
   k -3, kr 1.5, kw 16#8001, kt T#2s, ks SQRT(2.0). Worked by hand, the
   same at every tick:
   ABS(k): 3 (%QB0). MAX(k, 2): 2 (%QB1). LIMIT(0, k, 10): 0 (%QB2).
   SEL(k < 0, 1, 2): 2 (%QB3). MUX(1, 5, 6): 6 (%QB4).
   REAL_TO_INT(kr), 1.5 to the even one: 2 (%QB5); REAL_TO_INT(2.5): 2
   (%QB6); TRUNC_INT(kr): 1 (%QB7).
   SHL(kw, 1): 16#0002, 2 (%QB8). ROL(kw, 1): 16#0003, 3 (%QB9).
   ROR(kw, 17), by 1: 16#C000; shifted right by 12, 12 (%QB10).
   kt * 1.5 is T#3s: 1 (%QB11). kt / 3 is T#666ms: 1 (%QB12).
   kr ** 2, 2.25, times 4.0: 9 (%QB13). SQRT(2.0) times 10.0: 14
   (%QB14). 1.0 / 3.0 times 9.0: 3 (%QB15). ks * ks, 1.9999999, times
   50.0: 100 (%QB16). SQRT(2.0) > 1.0: TRUE (%QX17.0). SEL(ks > 1.0, 1,
   2): 2 (%QB18). lr : LREAL := EXP(LN(2.0)), times 50.0: 100 (%QB19).
   arr := [SQRT(4.0), SQRT(9.0)]: arr[1] + arr[2] is 5 (%QB20).
   The structure PT: x := ABS(-4), 4 (%QB21); y := SQRT(16.0), 4
   (%QB22). The TYPE RtT : REAL := SQRT(9.0): 3 (%QB23).
   The block F: inp := fk ** 2, fk 3.0: 9 (%QB24). The FUNCTION G: a :=
   SQRT(4.0) and loc := EXPT(2.0, 3): G() is 10 (%QB25), G(a := 1.0) 9
   (%QB26). The global gx := SQRT(INT_TO_REAL(g + 9)), g 7: 4 (%QB27).
   cv : DINT := INT_TO_DINT(k) * 1000, -3000, over 100: -30 (%QB28).
   u : USINT := INT_TO_USINT(ABS(k)): 3 (%QB29).
   A part of a constant array or structure is a constant: ka := [4,
   2(5)], k2 := [1, 2, 3, 4] of [1..2, 0..1], kp := (x := 6), kps :=
   [(x := 11), (x := 12, y := 2.5)], kr2 := [SQRT(4.0), 1.5].
   ka[2] + ka[k + 4], 5 + 4: 9 (%QB30). k2[2, 0]: 3 (%QB31). kp.x +
   kps[2].x: 18 (%QB32). kps[2].y * 2.0: 5 (%QB33). kp.y, its type's
   SQRT(16.0): 4 (%QB34). pf : PT := kps[2]: pf.x 12 (%QB35), pf.y
   times 2.0, 5 (%QB36). kr2[1] + kr2[2], 3.5, times 2.0: 7 (%QB37).
   ph := [ka[1], kp.x]: ph[1] + ph[2] is 10 (%QB38).
   reference-skip: the reference compiler takes no constant in an
   initial value (as constinit). *)
TYPE
  PT : STRUCT x : INT := ABS(-4); y : REAL := SQRT(16.0); END_STRUCT;
  RtT : REAL := SQRT(9.0);
END_TYPE
FUNCTION G : INT
  VAR_INPUT a : REAL := SQRT(4.0); END_VAR
  VAR loc : REAL := EXPT(2.0, 3); END_VAR
  G := REAL_TO_INT(a + loc);
END_FUNCTION
FUNCTION_BLOCK F
  VAR CONSTANT fk : REAL := 3.0; END_VAR
  VAR_INPUT inp : REAL := fk ** 2; END_VAR
  VAR_OUTPUT o : INT; END_VAR
  o := REAL_TO_INT(inp);
END_FUNCTION_BLOCK
CONFIGURATION c
  VAR_GLOBAL CONSTANT g : INT := 7; END_VAR
  VAR_GLOBAL gx : REAL := SQRT(INT_TO_REAL(g + 9)); END_VAR
  RESOURCE r ON x
    TASK t(INTERVAL := T#10ms, PRIORITY := 1);
    PROGRAM p WITH t : main;
  END_RESOURCE
END_CONFIGURATION
PROGRAM main
  VAR CONSTANT
    k : INT := -3;
    kr : REAL := 1.5;
    kw : WORD := 16#8001;
    kt : TIME := T#2s;
    ks : REAL := SQRT(2.0);
    ka : ARRAY [1..3] OF INT := [4, 2(5)];
    k2 : ARRAY [1..2, 0..1] OF INT := [1, 2, 3, 4];
    kp : PT := (x := 6);
    kps : ARRAY [1..2] OF PT := [(x := 11), (x := 12, y := 2.5)];
    kr2 : ARRAY [1..2] OF REAL := [SQRT(4.0), 1.5];
  END_VAR
  VAR_EXTERNAL gx : REAL; END_VAR
  VAR
    a : INT := ABS(k);
    b : INT := MAX(k, 2);
    c : INT := LIMIT(0, k, 10);
    d : INT := SEL(k < 0, 1, 2);
    e : INT := MUX(1, 5, 6);
    f1 : INT := REAL_TO_INT(kr);
    f2 : INT := REAL_TO_INT(2.5);
    f3 : INT := TRUNC_INT(kr);
    w1 : WORD := SHL(kw, 1);
    w2 : WORD := ROL(kw, 1);
    w3 : WORD := ROR(kw, 17);
    t1 : TIME := kt * 1.5;
    t2 : TIME := kt / 3;
    r1 : REAL := kr ** 2;
    r2 : REAL := SQRT(2.0);
    r3 : REAL := 1.0 / 3.0;
    r4 : REAL := ks * ks;
    bb : BOOL := SQRT(2.0) > 1.0;
    s1 : INT := SEL(ks > 1.0, 1, 2);
    lr : LREAL := EXP(LN(2.0));
    arr : ARRAY [1..2] OF REAL := [SQRT(4.0), SQRT(9.0)];
    p : PT;
    rt : RtT;
    fi : F;
    cv : DINT := INT_TO_DINT(k) * 1000;
    u : USINT := INT_TO_USINT(ABS(k));
    pa : INT := ka[2] + ka[k + 4];
    pb : INT := k2[2, 0];
    pc : INT := kp.x + kps[2].x;
    pd : REAL := kps[2].y * 2.0;
    pe : REAL := kp.y;
    pf : PT := kps[2];
    pg : REAL := kr2[1] + kr2[2];
    ph : ARRAY [1..2] OF INT := [ka[1], kp.x];
  END_VAR
  VAR
    q0 AT %QB0 : SINT;
    q1 AT %QB1 : SINT;
    q2 AT %QB2 : SINT;
    q3 AT %QB3 : SINT;
    q4 AT %QB4 : SINT;
    q5 AT %QB5 : SINT;
    q6 AT %QB6 : SINT;
    q7 AT %QB7 : SINT;
    q8 AT %QB8 : SINT;
    q9 AT %QB9 : SINT;
    q10 AT %QB10 : SINT;
    q11 AT %QB11 : SINT;
    q12 AT %QB12 : SINT;
    q13 AT %QB13 : SINT;
    q14 AT %QB14 : SINT;
    q15 AT %QB15 : SINT;
    q16 AT %QB16 : SINT;
    q17 AT %QX17.0 : BOOL;
    q18 AT %QB18 : SINT;
    q19 AT %QB19 : SINT;
    q20 AT %QB20 : SINT;
    q21 AT %QB21 : SINT;
    q22 AT %QB22 : SINT;
    q23 AT %QB23 : SINT;
    q24 AT %QB24 : SINT;
    q25 AT %QB25 : SINT;
    q26 AT %QB26 : SINT;
    q27 AT %QB27 : SINT;
    q28 AT %QB28 : SINT;
    q29 AT %QB29 : SINT;
    q30 AT %QB30 : SINT;
    q31 AT %QB31 : SINT;
    q32 AT %QB32 : SINT;
    q33 AT %QB33 : SINT;
    q34 AT %QB34 : SINT;
    q35 AT %QB35 : SINT;
    q36 AT %QB36 : SINT;
    q37 AT %QB37 : SINT;
    q38 AT %QB38 : SINT;
  END_VAR
  q0 := INT_TO_SINT(a);
  q1 := INT_TO_SINT(b);
  q2 := INT_TO_SINT(c);
  q3 := INT_TO_SINT(d);
  q4 := INT_TO_SINT(e);
  q5 := INT_TO_SINT(f1);
  q6 := INT_TO_SINT(f2);
  q7 := INT_TO_SINT(f3);
  q8 := WORD_TO_SINT(w1);
  q9 := WORD_TO_SINT(w2);
  q10 := WORD_TO_SINT(SHR(w3, 12));
  IF t1 = T#3s THEN
    q11 := 1;
  END_IF;
  IF t2 = T#666ms THEN
    q12 := 1;
  END_IF;
  q13 := REAL_TO_SINT(r1 * 4.0);
  q14 := REAL_TO_SINT(r2 * 10.0);
  q15 := REAL_TO_SINT(r3 * 9.0);
  q16 := REAL_TO_SINT(r4 * 50.0);
  q17 := bb;
  q18 := INT_TO_SINT(s1);
  q19 := LREAL_TO_SINT(lr * 50.0);
  q20 := REAL_TO_SINT(arr[1] + arr[2]);
  q21 := INT_TO_SINT(p.x);
  q22 := REAL_TO_SINT(p.y);
  q23 := REAL_TO_SINT(rt);
  fi();
  q24 := INT_TO_SINT(fi.o);
  q25 := INT_TO_SINT(G());
  q26 := INT_TO_SINT(G(a := 1.0));
  q27 := REAL_TO_SINT(gx);
  q28 := DINT_TO_SINT(cv / 100);
  q29 := USINT_TO_SINT(u);
  q30 := INT_TO_SINT(pa);
  q31 := INT_TO_SINT(pb);
  q32 := INT_TO_SINT(pc);
  q33 := REAL_TO_SINT(pd);
  q34 := REAL_TO_SINT(pe);
  q35 := INT_TO_SINT(pf.x);
  q36 := REAL_TO_SINT(pf.y * 2.0);
  q37 := REAL_TO_SINT(pg * 2.0);
  q38 := INT_TO_SINT(ph[1] + ph[2]);
END_PROGRAM

(* ---- constinit.st ---- *)
(* Initial values that are constant expressions (Ed.3 6.6.1.2.4,
   Figure 6): literals, CONSTANT variables and operators, worked out by
   the compiler - an integer one exactly, as the checker does it, a REAL
   one in single precision - for a variable, an array, a structure, a
   string, a block's and a FUNCTION's inputs and own variables.
   k 3, kr 1.5, kt T#2s, ks 'ab', kb TRUE; k2 := k + 1, 4; k3 := k2 * k,
   12; g, a global constant, 7. Worked by hand, the same at every tick:
   a := k * 2 + 1: 7 (%QB0). r := kr * 2.0: 3.0 (%QB1). r2 := kr / 4.0,
   0.375, times 8.0: 3 (%QB2). t := kt + T#500ms is T#2s500ms: 1 (%QB3).
   s := ks: LEN 2 (%QB4). b := NOT kb OR k > 2: TRUE (%QX5.0).
   arr : ARRAY [1..k] := [k, 2(k3)]: arr[3] 12 (%QB6). p := (x := k2, y
   := kr): p.x 4 (%QB7).
   The block FT: inp := fk + g, its constant 10 and the global 7: 17
   (%QB8). The FUNCTION G: a := c * 2 and loc := c + 1, c 5: G() 10 + 6,
   16 (%QB9); G(a := 1) 7 (%QB10).
   lvl : INT (0..10) := k: 3 (%QB11). m : MODE := run (%QB12 1).
   n := -k: -3 (%QB13). lr : LREAL := kr, times 2.0: 3 (%QB14).
   d : DINT := k3 * 10000, exactly 120000 though k3 is an INT: d / 10000
   is 12 (%QB15).
   A TYPE and a VAR_GLOBAL see the global constants directly: UT := g +
   1, 8 (%QB16), though the block HT has a constant g of its own, 1
   (%QB17); gx := g * 2: 14 (%QB18). A block's constant in its method:
   get's input a := mc, 4, and its x := mc + 1, 5: 9 (%QB19); in a
   block derived from it, v := mc * 3: 12 (%QB20).
   A constant of an enumeration, m2 := km, km run: 1 (%QB21). Bit
   strings: bb := 16#0F AND 16#3C, 16#0C: 12 (%QB22); bx := kx XOR
   16#05, kx 16#0F: 10 (%QB23). A named value, nv := hi + 1: 6 (%QB24).
   reference-skip: the reference compiler takes no constant in an
   initial value or a bound (as flexarrays). *)
TYPE
  PT : STRUCT x : INT; y : REAL; END_STRUCT;
  MODE : (idle, run);
  UT : INT := g + 1;
  LV : INT (lo := 1, hi := 5);
END_TYPE
FUNCTION_BLOCK HT
  VAR CONSTANT g : INT := 1; END_VAR
  VAR_OUTPUT u : UT; own : INT := g; END_VAR
END_FUNCTION_BLOCK
FUNCTION_BLOCK MT
  VAR CONSTANT mc : INT := 4; END_VAR
  METHOD PUBLIC get : INT
    VAR_INPUT a : INT := mc; END_VAR
    VAR x : INT := mc + 1; END_VAR
    get := a + x;
  END_METHOD
END_FUNCTION_BLOCK
FUNCTION_BLOCK DTB EXTENDS MT
  VAR_OUTPUT v : INT := mc * 3; END_VAR
END_FUNCTION_BLOCK
FUNCTION_BLOCK FT
  VAR CONSTANT fk : INT := 10; END_VAR
  VAR_EXTERNAL CONSTANT g : INT; END_VAR
  VAR_INPUT inp : INT := fk + g; END_VAR
  VAR_OUTPUT o : INT; END_VAR
  o := inp;
END_FUNCTION_BLOCK
FUNCTION G : INT
  VAR CONSTANT c : INT := 5; END_VAR
  VAR_INPUT a : INT := c * 2; END_VAR
  VAR loc : INT := c + 1; END_VAR
  G := a + loc;
END_FUNCTION
CONFIGURATION c
  VAR_GLOBAL CONSTANT g : INT := 7; END_VAR
  VAR_GLOBAL gx : INT := g * 2; END_VAR
  RESOURCE r ON PLC
    TASK t(INTERVAL := T#10ms, PRIORITY := 1);
    PROGRAM p WITH t : main;
  END_RESOURCE
END_CONFIGURATION
PROGRAM main
  VAR CONSTANT
    k : INT := 3;
    kr : REAL := 1.5;
    kt : TIME := T#2s;
    ks : STRING := 'ab';
    kb : BOOL := TRUE;
    k2 : INT := k + 1;
    k3 : INT := k2 * k;
    km : MODE := run;
    kx : BYTE := 16#0F;
  END_VAR
  VAR_EXTERNAL gx : INT; END_VAR
  VAR
    a : INT := k * 2 + 1;
    r : REAL := kr * 2.0;
    r2 : REAL := kr / 4.0;
    t : TIME := kt + T#500ms;
    s : STRING := ks;
    b : BOOL := NOT kb OR k > 2;
    arr : ARRAY [1..k] OF INT := [k, 2(k3)];
    p : PT := (x := k2, y := kr);
    f : FT;
    lvl : INT (0..10) := k;
    m : MODE := run;
    n : INT := -k;
    lr : LREAL := kr;
    d : DINT := k3 * 10000;
    h : HT;
    mi : MT;
    di : DTB;
    m2 : MODE := km;
    bb : BYTE := 16#0F AND 16#3C;
    bx : BYTE := kx XOR 16#05;
    nv : INT := hi + 1;
  END_VAR
  VAR
    q0 AT %QB0 : SINT;
    q1 AT %QB1 : SINT;
    q2 AT %QB2 : SINT;
    q3 AT %QB3 : SINT;
    q4 AT %QB4 : SINT;
    q5 AT %QX5.0 : BOOL;
    q6 AT %QB6 : SINT;
    q7 AT %QB7 : SINT;
    q8 AT %QB8 : SINT;
    q9 AT %QB9 : SINT;
    q10 AT %QB10 : SINT;
    q11 AT %QB11 : SINT;
    q12 AT %QB12 : SINT;
    q13 AT %QB13 : SINT;
    q14 AT %QB14 : SINT;
    q15 AT %QB15 : SINT;
    q16 AT %QB16 : SINT;
    q17 AT %QB17 : SINT;
    q18 AT %QB18 : SINT;
    q19 AT %QB19 : SINT;
    q20 AT %QB20 : SINT;
    q21 AT %QB21 : SINT;
    q22 AT %QB22 : SINT;
    q23 AT %QB23 : SINT;
    q24 AT %QB24 : SINT;
  END_VAR
  q0 := INT_TO_SINT(a);
  q1 := REAL_TO_SINT(r);
  q2 := REAL_TO_SINT(r2 * 8.0);
  IF t = T#2s500ms THEN
    q3 := 1;
  END_IF;
  q4 := INT_TO_SINT(LEN(s));
  q5 := b;
  q6 := INT_TO_SINT(arr[3]);
  q7 := INT_TO_SINT(p.x);
  f();
  q8 := INT_TO_SINT(f.o);
  q9 := INT_TO_SINT(G());
  q10 := INT_TO_SINT(G(a := 1));
  q11 := INT_TO_SINT(lvl);
  IF m = run THEN
    q12 := 1;
  END_IF;
  q13 := INT_TO_SINT(n);
  q14 := LREAL_TO_SINT(lr * 2.0);
  q15 := DINT_TO_SINT(d / 10000);
  q16 := INT_TO_SINT(h.u);
  q17 := INT_TO_SINT(h.own);
  q18 := INT_TO_SINT(gx);
  q19 := INT_TO_SINT(mi.get());
  q20 := INT_TO_SINT(di.v);
  IF m2 = run THEN
    q21 := 1;
  END_IF;
  q22 := BYTE_TO_SINT(bb);
  q23 := BYTE_TO_SINT(bx);
  q24 := INT_TO_SINT(nv);
END_PROGRAM

(* ---- debugsteps.st ---- *)
(* A debug build (docs/c-output.md §10): the hook before each statement
   as it runs, with its POU, line and instance. A block's two
   instances say which is running; a FUNCTION has none; IF and FOR run
   their own line, then their statements'. Worked by hand, one tick:

   main 27 (c1()), then cnt's 21 and 22 in R.P.C1 (n 1, not > 100);
   main 28, then 21 and 22 in R.P.C2; main 29 (q := twice(c1.n)), then
   twice's 17, no instance; main 30 (the IF: c1.n is 1), then 31; main
   33 (the FOR), then its body, 34, for i 1 and for i 2, the FOR's 33
   before each later test (i 2, then i 3, which ends it); main 36 (the
   IF, s2 3 not > 10), 38 (its ELSIF, s2 = 3), 39; main 41 (the WHILE,
   i 3 > 2), 42, i 2, 41 again (not > 2: done); main 44 (the REPEAT),
   45, i 1, then its UNTIL 46 (1 < 2: done). q is 2 + 1 + 10 (Q0 0d
   00). *)
FUNCTION twice : INT
  VAR_INPUT x : INT; END_VAR
  twice := x * 2;
END_FUNCTION
FUNCTION_BLOCK cnt
  VAR_OUTPUT n : INT; END_VAR
  n := n + 1;
  IF n > 100 THEN n := 0; END_IF;
END_FUNCTION_BLOCK
PROGRAM main
  VAR c1, c2 : cnt; i, s2 : INT; END_VAR
  VAR q AT %QW0 : INT; END_VAR
  c1();
  c2();
  q := twice(c1.n);
  IF c1.n = 1 THEN
    q := q + 1;
  END_IF;
  FOR i := 1 TO 2 DO
    s2 := s2 + i;
  END_FOR;
  IF s2 > 10 THEN
    q := 0;
  ELSIF s2 = 3 THEN
    q := q + 10;
  END_IF;
  WHILE i > 2 DO
    i := i - 1;
  END_WHILE;
  REPEAT
    i := i - 1;
  UNTIL i < 2
  END_REPEAT;
END_PROGRAM
CONFIGURATION c RESOURCE r ON PLC TASK t(INTERVAL := T#10ms, PRIORITY := 1); PROGRAM p WITH t : main; END_RESOURCE END_CONFIGURATION

(* ---- directwrite.st ---- *)
(* Directly represented variables written in a body (Ed.3 6.5.5,
   deprecated: W0002): assigned, a block's output and ENO taken into
   one, one given to a FUNCTION's and a block's in-out. %IX1.0 TRUE,
   %IW2 16#1234, %IX0.2 TRUE from tick 0. Worked by hand:

   tick 0: %QX1.0 := %IX1.0, 1 (Q1 01); %QW2 := %IW2 (Q2 34 12); the
   TON's Q into %QX0.3, not yet; fo's ENO into %QX0.0, TRUE (Q0 01);
   setb sets bit 0 of %MW4 through its in-out (M4 01); the block sets
   bit 8 of %MW6 (M7 01); w counts, 1 (Q4 01). The program io, its
   in-out connected to %MW8 in the CONFIGURATION, shifts a 1 into it:
   1 (M8 01).
   tick 1: w 2, %MW8 3. tick 2: w 3, %MW8 7, and the TON is done after
   20 ms: %QX0.3 (Q0 09).
   reference-skip: the reference compiler's C writes no direct address
   in a body. *)
FUNCTION setb : WORD
  VAR_IN_OUT x : WORD; END_VAR
  x := x OR 16#0001;
  setb := x;
END_FUNCTION
FUNCTION fo : INT
  VAR_INPUT x : INT; END_VAR
  fo := x;
END_FUNCTION
FUNCTION_BLOCK blk
  VAR_IN_OUT x : WORD; END_VAR
  x := x OR 16#0100;
END_FUNCTION_BLOCK
PROGRAM main
  VAR t : TON; w : USINT; k : INT; b : blk; r : WORD; END_VAR
  %QX1.0 := %IX1.0;
  %QW2 := %IW2;
  t(IN := %IX0.2, PT := T#20ms, Q => %QX0.3);
  k := fo(EN := %IX0.2, x := 1, ENO => %QX0.0);
  r := setb(%MW4);
  b(x := %MW6);
  w := w + 1;
  %QB4 := USINT_TO_BYTE(w);
END_PROGRAM
PROGRAM io
  VAR_IN_OUT n : WORD; END_VAR
  n := ROL(n, 1) OR 16#0001;
END_PROGRAM
CONFIGURATION c
  RESOURCE r ON PLC
    TASK t(INTERVAL := T#10ms, PRIORITY := 1);
    PROGRAM p WITH t : main;
    PROGRAM p2 WITH t : io(n := %MW8);
  END_RESOURCE
END_CONFIGURATION

(* ---- edgeinputs.st ---- *)
(* R_EDGE and F_EDGE inputs of a FUNCTION_BLOCK and a PROGRAM (Ed.3
   6.6.3.2 rule 13, Table 40 6a): an implicit R_TRIG or F_TRIG in the
   instance; the body sees its Q. The input %IX0.0 is FALSE at tick 0,
   TRUE at 1 and 2, FALSE at 3, TRUE at 4. Worked by hand, ticks 0..4:
   ET counts clk's rising edges in n: 0 1 1 1 2 (%QB0); fall's falling
   ones in m: an F_TRIG first called with CLK FALSE gives Q TRUE once
   (Table 44: M starts FALSE), so 1 1 1 2 2 (%QB1).
   The PROGRAM's own x, connected to %IX0.0, counted in p: 0 1 1 1 2
   (%QB2). Read from outside, e.clk is what was given, not the edge:
   0 1 1 0 1 (%QX3.0).
   reference-skip: R_EDGE and F_EDGE: the reference compiler does not
   support them. *)
FUNCTION_BLOCK ET
  VAR_INPUT clk : BOOL R_EDGE; fall : BOOL F_EDGE; END_VAR
  VAR_OUTPUT n : INT; m : INT; END_VAR
  IF clk THEN
    n := n + 1;
  END_IF;
  IF fall THEN
    m := m + 1;
  END_IF;
END_FUNCTION_BLOCK
PROGRAM main
  VAR_INPUT x : BOOL R_EDGE; END_VAR
  VAR
    e : ET;
    p : INT;
  END_VAR
  VAR
    i AT %IX0.0 : BOOL;
    q0 AT %QB0 : SINT;
    q1 AT %QB1 : SINT;
    q2 AT %QB2 : SINT;
    q3 AT %QX3.0 : BOOL;
  END_VAR
  e(clk := i, fall := i);
  q0 := INT_TO_SINT(e.n);
  q1 := INT_TO_SINT(e.m);
  IF x THEN
    p := p + 1;
  END_IF;
  q2 := INT_TO_SINT(p);
  q3 := e.clk;
END_PROGRAM

CONFIGURATION c
  RESOURCE r ON x
    TASK t(INTERVAL := T#10ms, PRIORITY := 1);
    PROGRAM pr WITH t : main(x := %IX0.0);
  END_RESOURCE
END_CONFIGURATION

(* ---- endiancorners.st ---- *)
(* The endianness functions (Ed.3 6.6.2.5.13) of what holds more than
   data: a structure holding an instance, a structure with `*`
   components, and ARRAY[*]. Worked by hand, on a little-endian target:
   tick 0 (%ID0 16#01020304):
   x.c, a CTU in Box, counts once: CV 1. y := TO_BIG_ENDIAN(x): y.w
   16#0A0B0C0D reversed, MD32 0a 0b 0c 0d; y.c copied as it is, an
   instance being no data type's value: CV 1 (MW36 01 00).
   a.out := 16#CAFEBABE at %QD0 (be ba fe ca); a.k := 16#1234. b :=
   TO_BIG_ENDIAN(a): each `*` part converted in a buffer of its own, so
   a's addresses are not written: Q0 stays be ba fe ca, b.out at %QD4 is
   ca fe ba be; b.raw at %ID4 is a.raw reversed; bk := b.k, 16#3412
   (MW40 12 34). braw := b.raw reads it back: 16#04030201 (MD42 01 02
   03 04).
   s(a := p, b := q, m := g, n := h): q := TO_BIG_ENDIAN(p) stored, then
   converted where it is: MD8 11 22 33 44 55 66 77 88; h :=
   FROM_BIG_ENDIAN(g), each INT reversed: MW24 01 02 03 04 05 06 07 08;
   r := TO_LITTLE_ENDIAN(z) (z of fixed bounds into an ARRAY[*]) as it
   is: MD46 78 56 34 12.
   tick 1: the CTU's CU stays TRUE: CV 1 still; the rest as tick 0.
   reference-skip: the reference compiler (Ed.2) has neither the
   endianness functions nor ARRAY[*], and generates nothing for
   VAR_CONFIG. *)
TYPE
  Box : STRUCT c : CTU; w : DWORD; END_STRUCT;
  IoW : STRUCT raw AT %I* : DWORD; out AT %Q* : DWORD; k : WORD; END_STRUCT;
END_TYPE
FUNCTION_BLOCK Swap
  VAR_IN_OUT a, b, r : ARRAY[*] OF DWORD; m, n : ARRAY[*, *] OF INT; END_VAR
  VAR z : ARRAY[0..0] OF DWORD := [16#12345678]; END_VAR
  b := TO_BIG_ENDIAN(a);
  n := FROM_BIG_ENDIAN(m);
  r := TO_LITTLE_ENDIAN(z);
END_FUNCTION_BLOCK
PROGRAM line
  VAR x, y : Box; a, b : IoW; s : Swap; END_VAR
  VAR
    p AT %MD0 : ARRAY[0..1] OF DWORD := [16#11223344, 16#55667788];
    q AT %MD8 : ARRAY[0..1] OF DWORD;
    g AT %MW16 : ARRAY[0..1, 0..1] OF INT := [16#0102, 16#0304, 16#0506, 16#0708];
    h AT %MW24 : ARRAY[0..1, 0..1] OF INT;
    yw AT %MD32 : DWORD;
    ycv AT %MW36 : INT;
    bk AT %MW40 : WORD;
    braw AT %MD42 : DWORD;
    zr AT %MD46 : ARRAY[0..0] OF DWORD;
  END_VAR
  x.c(CU := TRUE, PV := 5);
  x.w := 16#0A0B0C0D;
  y := TO_BIG_ENDIAN(x);
  yw := y.w;
  ycv := y.c.CV;
  a.out := 16#CAFEBABE;
  a.k := 16#1234;
  b := TO_BIG_ENDIAN(a);
  bk := b.k;
  braw := b.raw;
  s(a := p, b := q, m := g, n := h, r := zr);
END_PROGRAM
CONFIGURATION plant
  RESOURCE cpu ON PLC
    TASK fast (INTERVAL := T#10ms, PRIORITY := 1);
    PROGRAM main WITH fast : line;
  END_RESOURCE
  VAR_CONFIG
    cpu.main.a.raw AT %ID0 : DWORD;
    cpu.main.a.out AT %QD0 : DWORD;
    cpu.main.b.raw AT %ID4 : DWORD;
    cpu.main.b.out AT %QD4 : DWORD;
  END_VAR
END_CONFIGURATION
